PROGRAM OtherDevice_外部機器
VAR
    FH_M : BOOL;
    GT2_M : BOOL;
    IAI_M : BOOL;
    HMI_M : BOOL;
    FH_A_ST1_M : ARRAY[0..99] OF Bool;  (* [1] ST1 FH測定中; [5] ST1 測定完了 *)
    FH_A_ST1_OK : BOOL;  (* ST1 OK判定 *)
    FH_A_ST1_NG : BOOL;  (* ST1 NG 判定 *)
    FH_A_ST1_TON : ARRAY[0..99] OF TON;
    FH_A_ST1_TOF : ARRAY[0..99] OF TOF;
    ４ : UINT;
    ConvWordIndex : INT;  (* ワード処理ループの添字。（2台を順番に処理する作業用。運転指令は入れない） *)
    ConvAxisIndex : INT;  (* 軸処理ループの添字1～6。（2台を順番に処理する作業用。運転指令は入れない） *)
    ConvBase : INT;  (* 軸データの先頭添字8/16/24/32/40/48。（2台を順番に処理する作業用。運転指令は入れない） *)
    ConvDWord : DWORD;  (* 32bitの分割・結合に使うビット列。（2台を順番に処理する作業用。運転指令は入れない） *)
    ConvPos : DINT;  (* 0.01mm単位の符号付き目標位置。（2台を順番に処理する作業用。運転指令は入れない） *)
    ConvBand : UDINT;  (* 0.01mm単位の非負位置決め幅（内部推奨型）。（2台を順番に処理する作業用。運転指令は入れない） *)
    ConvSpeed : UINT;  (* 速度の送信整数。（2台を順番に処理する作業用。運転指令は入れない） *)
    ConvAccDec : UINT;  (* 加減速度の送信整数。（2台を順番に処理する作業用。運転指令は入れない） *)
    ConvPush : UINT;  (* 押付け電流制限の送信整数。（2台を順番に処理する作業用。運転指令は入れない） *)
    ConvScaled : LREAL;  (* 単位換算の作業値。（2台を順番に処理する作業用。運転指令は入れない） *)
    ConvWord : WORD;  (* バイト交換の作業ワード。（2台を順番に処理する作業用。運転指令は入れない） *)
    ConvUnitOK : BOOL;  (* 速度単位が1.0または0.1であること。（2台を順番に処理する作業用。運転指令は入れない） *)
END_VAR
VAR_EXTERNAL
    HMI_MessageNo : ARRAY[0..9] OF UINT;
    HMI_Message : ARRAY[0..9] OF String[256];
    HMI_Language : BOOL;
    FH_Line0_Trigger_Ready_1 : BOOL;
    FH_Line0_Trigger_1 : BOOL;
    M9999 : BOOL;
    FH_Line0_Busy_1 : BOOL;
    FH_Line0_Result_Notification_1 : BOOL;
    FH_Line0_DINT_Result_Data_0_1 : DINT;
    FH_Line0_DINT_Result_Data_1_1 : DINT;
    FH_Line0_DINT_Result_Data_2_1 : DINT;
    FH_Line0_Command_Code_1 : DWORD;
    FH_Line0_Command_Request_1 : BOOL;
    FH_Line0_Command_Completion_1 : BOOL;
    MdlChg : BOOL;  (* 機種切替：ON【GA120】 OFF【GA90】 *)
    FH_Line0_Error_Status_1 : BOOL;
    FH_5552_10_A_Auto : BOOL;  (* ST1 FH測定開始 *)
    FH_A_ST1_Manual : BOOL;  (* ST1 *)
    Pause : ARRAY[0..99] OF Bool;
    FH_A_ST1_Done : BOOL;  (* ST1 画像検査完了 *)
    Station_A_Data : ARRAY[0..8] OF sData;
    DLEP1_OUT : ARRAY[0..79] OF BOOL;
    DLEP2_OUT : ARRAY[0..79] OF BOOL;
    DLEP1_IN : ARRAY[0..167] OF byte;
    DLEP2_IN : ARRAY[0..167] OF byte;
    DLEP2_IN_Error : BOOL;  (* B(右側)センサエラー *)
    DLEP1_IN_Error : BOOL;  (* A(右側)センサエラー *)
    GT2_A_CurrentVal : INT;  (* A(左側) 測定値 *)
    GT2_B_CurrentVal : INT;  (* B(右側) 測定値 *)
    Hgt_A_Ins_Data : LREAL;  (* A測定データに変換 *)
    Hgt_B_Ins_Data : LREAL;
    Hgt_A_ComputedValueData : LREAL;  (* A測定データ+13.000mm 算定データ *)
    Hgt_B_ComputedValueData : LREAL;  (* B測定データ+13.000mm 算定データ *)
    E001_In_IN00_2004_01 : UINT;  (* RCON1（Node1） RCON→PLC 【IN00】共通 ゲートウェイ状態信号0 *)
    E001_In_IN01_2004_02 : UINT;  (* RCON1（Node1） RCON→PLC 【IN01】共通 ゲートウェイ状態信号1（軸No.0～15リンク状態） *)
    E001_In_IN02_2004_03 : UINT;  (* RCON1（Node1） RCON→PLC 【IN02】共通 電源ユニット状態信号0 *)
    E001_In_IN03_2004_04 : UINT;  (* RCON1（Node1） RCON→PLC 【IN03】共通 電源ユニット状態信号1 *)
    E001_In_IN04_2004_05 : UINT;  (* RCON1（Node1） RCON→PLC 【IN04】共通 電源ユニット状態信号2 *)
    E001_In_IN05_2004_06 : UINT;  (* RCON1（Node1） RCON→PLC 【IN05】共通 電源ユニット状態信号3 *)
    E001_In_IN06_2004_07 : UINT;  (* RCON1（Node1） RCON→PLC 【IN06】共通 電源ユニット状態信号4／軽故障メンテナンス（設定依存） *)
    E001_In_IN07_2004_08 : UINT;  (* RCON1（Node1） RCON→PLC 【IN07】共通 共通予約領域（使用禁止・占有あり） *)
    E001_In_IN08_2004_09 : UINT;  (* RCON1（Node1） RCON→PLC 【IN08】1軸目（No.0） 現在位置 下位ワード *)
    E001_In_IN09_2004_0A : UINT;  (* RCON1（Node1） RCON→PLC 【IN09】1軸目（No.0） 現在位置 上位ワード *)
    E001_In_IN10_2004_0B : UINT;  (* RCON1（Node1） RCON→PLC 【IN10】1軸目（No.0） 現在電流 下位ワード（PCは指令電流） *)
    E001_In_IN11_2004_0C : UINT;  (* RCON1（Node1） RCON→PLC 【IN11】1軸目（No.0） 現在電流 上位ワード（PCは指令電流） *)
    E001_In_IN12_2004_0D : UINT;  (* RCON1（Node1） RCON→PLC 【IN12】1軸目（No.0） 現在速度（負方向は2の補数） *)
    E001_In_IN13_2004_0E : UINT;  (* RCON1（Node1） RCON→PLC 【IN13】1軸目（No.0） 予約領域（使用禁止） *)
    E001_In_IN14_2004_0F : UINT;  (* RCON1（Node1） RCON→PLC 【IN14】1軸目（No.0） アラームコード（簡易コードではない） *)
    E001_In_IN15_2004_10 : UINT;  (* RCON1（Node1） RCON→PLC 【IN15】1軸目（No.0） 軸状態信号（PEND・SV等） *)
    E001_In_IN16_2004_11 : UINT;  (* RCON1（Node1） RCON→PLC 【IN16】2軸目（No.1） 現在位置 下位ワード *)
    E001_In_IN17_2004_12 : UINT;  (* RCON1（Node1） RCON→PLC 【IN17】2軸目（No.1） 現在位置 上位ワード *)
    E001_In_IN18_2004_13 : UINT;  (* RCON1（Node1） RCON→PLC 【IN18】2軸目（No.1） 現在電流 下位ワード（PCは指令電流） *)
    E001_In_IN19_2004_14 : UINT;  (* RCON1（Node1） RCON→PLC 【IN19】2軸目（No.1） 現在電流 上位ワード（PCは指令電流） *)
    E001_In_IN20_2004_15 : UINT;  (* RCON1（Node1） RCON→PLC 【IN20】2軸目（No.1） 現在速度（負方向は2の補数） *)
    E001_In_IN21_2004_16 : UINT;  (* RCON1（Node1） RCON→PLC 【IN21】2軸目（No.1） 予約領域（使用禁止） *)
    E001_In_IN22_2004_17 : UINT;  (* RCON1（Node1） RCON→PLC 【IN22】2軸目（No.1） アラームコード（簡易コードではない） *)
    E001_In_IN23_2004_18 : UINT;  (* RCON1（Node1） RCON→PLC 【IN23】2軸目（No.1） 軸状態信号（PEND・SV等） *)
    E001_In_IN24_2004_19 : UINT;  (* RCON1（Node1） RCON→PLC 【IN24】3軸目（No.2） 現在位置 下位ワード *)
    E001_In_IN25_2004_1A : UINT;  (* RCON1（Node1） RCON→PLC 【IN25】3軸目（No.2） 現在位置 上位ワード *)
    E001_In_IN26_2004_1B : UINT;  (* RCON1（Node1） RCON→PLC 【IN26】3軸目（No.2） 現在電流 下位ワード（PCは指令電流） *)
    E001_In_IN27_2004_1C : UINT;  (* RCON1（Node1） RCON→PLC 【IN27】3軸目（No.2） 現在電流 上位ワード（PCは指令電流） *)
    E001_In_IN28_2004_1D : UINT;  (* RCON1（Node1） RCON→PLC 【IN28】3軸目（No.2） 現在速度（負方向は2の補数） *)
    E001_In_IN29_2004_1E : UINT;  (* RCON1（Node1） RCON→PLC 【IN29】3軸目（No.2） 予約領域（使用禁止） *)
    E001_In_IN30_2004_1F : UINT;  (* RCON1（Node1） RCON→PLC 【IN30】3軸目（No.2） アラームコード（簡易コードではない） *)
    E001_In_IN31_2004_20 : UINT;  (* RCON1（Node1） RCON→PLC 【IN31】3軸目（No.2） 軸状態信号（PEND・SV等） *)
    E001_In_IN32_2004_21 : UINT;  (* RCON1（Node1） RCON→PLC 【IN32】4軸目（No.3） 現在位置 下位ワード *)
    E001_In_IN33_2004_22 : UINT;  (* RCON1（Node1） RCON→PLC 【IN33】4軸目（No.3） 現在位置 上位ワード *)
    E001_In_IN34_2004_23 : UINT;  (* RCON1（Node1） RCON→PLC 【IN34】4軸目（No.3） 現在電流 下位ワード（PCは指令電流） *)
    E001_In_IN35_2004_24 : UINT;  (* RCON1（Node1） RCON→PLC 【IN35】4軸目（No.3） 現在電流 上位ワード（PCは指令電流） *)
    E001_In_IN36_2004_25 : UINT;  (* RCON1（Node1） RCON→PLC 【IN36】4軸目（No.3） 現在速度（負方向は2の補数） *)
    E001_In_IN37_2004_26 : UINT;  (* RCON1（Node1） RCON→PLC 【IN37】4軸目（No.3） 予約領域（使用禁止） *)
    E001_In_IN38_2004_27 : UINT;  (* RCON1（Node1） RCON→PLC 【IN38】4軸目（No.3） アラームコード（簡易コードではない） *)
    E001_In_IN39_2004_28 : UINT;  (* RCON1（Node1） RCON→PLC 【IN39】4軸目（No.3） 軸状態信号（PEND・SV等） *)
    E001_In_IN40_2004_29 : UINT;  (* RCON1（Node1） RCON→PLC 【IN40】5軸目（No.4） 現在位置 下位ワード *)
    E001_In_IN41_2004_2A : UINT;  (* RCON1（Node1） RCON→PLC 【IN41】5軸目（No.4） 現在位置 上位ワード *)
    E001_In_IN42_2004_2B : UINT;  (* RCON1（Node1） RCON→PLC 【IN42】5軸目（No.4） 現在電流 下位ワード（PCは指令電流） *)
    E001_In_IN43_2004_2C : UINT;  (* RCON1（Node1） RCON→PLC 【IN43】5軸目（No.4） 現在電流 上位ワード（PCは指令電流） *)
    E001_In_IN44_2004_2D : UINT;  (* RCON1（Node1） RCON→PLC 【IN44】5軸目（No.4） 現在速度（負方向は2の補数） *)
    E001_In_IN45_2004_2E : UINT;  (* RCON1（Node1） RCON→PLC 【IN45】5軸目（No.4） 予約領域（使用禁止） *)
    E001_In_IN46_2004_2F : UINT;  (* RCON1（Node1） RCON→PLC 【IN46】5軸目（No.4） アラームコード（簡易コードではない） *)
    E001_In_IN47_2004_30 : UINT;  (* RCON1（Node1） RCON→PLC 【IN47】5軸目（No.4） 軸状態信号（PEND・SV等） *)
    E001_In_IN48_2004_31 : UINT;  (* RCON1（Node1） RCON→PLC 【IN48】6軸目（No.5） 現在位置 下位ワード *)
    E001_In_IN49_2004_32 : UINT;  (* RCON1（Node1） RCON→PLC 【IN49】6軸目（No.5） 現在位置 上位ワード *)
    E001_In_IN50_2004_33 : UINT;  (* RCON1（Node1） RCON→PLC 【IN50】6軸目（No.5） 現在電流 下位ワード（PCは指令電流） *)
    E001_In_IN51_2004_34 : UINT;  (* RCON1（Node1） RCON→PLC 【IN51】6軸目（No.5） 現在電流 上位ワード（PCは指令電流） *)
    E001_In_IN52_2004_35 : UINT;  (* RCON1（Node1） RCON→PLC 【IN52】6軸目（No.5） 現在速度（負方向は2の補数） *)
    E001_In_IN53_2004_36 : UINT;  (* RCON1（Node1） RCON→PLC 【IN53】6軸目（No.5） 予約領域（使用禁止） *)
    E001_In_IN54_2004_37 : UINT;  (* RCON1（Node1） RCON→PLC 【IN54】6軸目（No.5） アラームコード（簡易コードではない） *)
    E001_In_IN55_2004_38 : UINT;  (* RCON1（Node1） RCON→PLC 【IN55】6軸目（No.5） 軸状態信号（PEND・SV等） *)
    E001_In_IN56_2004_39 : UINT;  (* RCON1（Node1） 【IN56】用途未確認領域。今回の軸データ変換では未使用。 *)
    E001_In_IN57_2004_3A : UINT;  (* RCON1（Node1） 【IN57】用途未確認領域。今回の軸データ変換では未使用。 *)
    E001_In_IN58_2004_3B : UINT;  (* RCON1（Node1） 【IN58】用途未確認領域。今回の軸データ変換では未使用。 *)
    E001_In_IN59_2004_3C : UINT;  (* RCON1（Node1） 【IN59】用途未確認領域。今回の軸データ変換では未使用。 *)
    E001_In_IN60_2004_3D : UINT;  (* RCON1（Node1） 【IN60】用途未確認領域。今回の軸データ変換では未使用。 *)
    E001_In_IN61_2004_3E : UINT;  (* RCON1（Node1） 【IN61】用途未確認領域。今回の軸データ変換では未使用。 *)
    E001_In_IN62_2004_3F : UINT;  (* RCON1（Node1） 【IN62】用途未確認領域。今回の軸データ変換では未使用。 *)
    E001_In_IN63_2004_40 : UINT;  (* RCON1（Node1） 【IN63】用途未確認領域。今回の軸データ変換では未使用。 *)
    E001_In_IN64_2004_41 : UINT;  (* RCON1（Node1） 【IN64】用途未確認領域。今回の軸データ変換では未使用。 *)
    E001_In_IN65_2004_42 : UINT;  (* RCON1（Node1） 【IN65】用途未確認領域。今回の軸データ変換では未使用。 *)
    E001_In_IN66_2004_43 : UINT;  (* RCON1（Node1） 【IN66】用途未確認領域。今回の軸データ変換では未使用。 *)
    E001_In_IN67_2004_44 : UINT;  (* RCON1（Node1） 【IN67】用途未確認領域。今回の軸データ変換では未使用。 *)
    E001_In_IN68_2004_45 : UINT;  (* RCON1（Node1） 【IN68】用途未確認領域。今回の軸データ変換では未使用。 *)
    E001_In_IN69_2004_46 : UINT;  (* RCON1（Node1） 【IN69】用途未確認領域。今回の軸データ変換では未使用。 *)
    E001_In_IN70_2004_47 : UINT;  (* RCON1（Node1） 【IN70】用途未確認領域。今回の軸データ変換では未使用。 *)
    E001_In_IN71_2004_48 : UINT;  (* RCON1（Node1） 【IN71】用途未確認領域。今回の軸データ変換では未使用。 *)
    E001_Out_OUT00_2003_01 : UINT;  (* RCON1（Node1） PLC→RCON 【OUT00】共通 ゲートウェイ制御信号0（MON等） *)
    E001_Out_OUT08_2003_09 : UINT;  (* RCON1（Node1） PLC→RCON 【OUT08】1軸目（No.0） 目標位置 下位ワード *)
    E001_Out_OUT09_2003_0A : UINT;  (* RCON1（Node1） PLC→RCON 【OUT09】1軸目（No.0） 目標位置 上位ワード *)
    E001_Out_OUT10_2003_0B : UINT;  (* RCON1（Node1） PLC→RCON 【OUT10】1軸目（No.0） 位置決め幅 下位ワード *)
    E001_Out_OUT11_2003_0C : UINT;  (* RCON1（Node1） PLC→RCON 【OUT11】1軸目（No.0） 位置決め幅 上位ワード *)
    E001_Out_OUT12_2003_0D : UINT;  (* RCON1（Node1） PLC→RCON 【OUT12】1軸目（No.0） 速度指令 *)
    E001_Out_OUT13_2003_0E : UINT;  (* RCON1（Node1） PLC→RCON 【OUT13】1軸目（No.0） 加減速度指令（加速・減速共通） *)
    E001_Out_OUT14_2003_0F : UINT;  (* RCON1（Node1） PLC→RCON 【OUT14】1軸目（No.0） 押付け電流制限値 *)
    E001_Out_OUT15_2003_10 : UINT;  (* RCON1（Node1） PLC→RCON 【OUT15】1軸目（No.0） 軸制御信号（DSTR・SON等） *)
    E001_Out_OUT16_2003_11 : UINT;  (* RCON1（Node1） PLC→RCON 【OUT16】2軸目（No.1） 目標位置 下位ワード *)
    E001_Out_OUT17_2003_12 : UINT;  (* RCON1（Node1） PLC→RCON 【OUT17】2軸目（No.1） 目標位置 上位ワード *)
    E001_Out_OUT18_2003_13 : UINT;  (* RCON1（Node1） PLC→RCON 【OUT18】2軸目（No.1） 位置決め幅 下位ワード *)
    E001_Out_OUT19_2003_14 : UINT;  (* RCON1（Node1） PLC→RCON 【OUT19】2軸目（No.1） 位置決め幅 上位ワード *)
    E001_Out_OUT20_2003_15 : UINT;  (* RCON1（Node1） PLC→RCON 【OUT20】2軸目（No.1） 速度指令 *)
    E001_Out_OUT21_2003_16 : UINT;  (* RCON1（Node1） PLC→RCON 【OUT21】2軸目（No.1） 加減速度指令（加速・減速共通） *)
    E001_Out_OUT22_2003_17 : UINT;  (* RCON1（Node1） PLC→RCON 【OUT22】2軸目（No.1） 押付け電流制限値 *)
    E001_Out_OUT23_2003_18 : UINT;  (* RCON1（Node1） PLC→RCON 【OUT23】2軸目（No.1） 軸制御信号（DSTR・SON等） *)
    E001_Out_OUT24_2003_19 : UINT;  (* RCON1（Node1） PLC→RCON 【OUT24】3軸目（No.2） 目標位置 下位ワード *)
    E001_Out_OUT25_2003_1A : UINT;  (* RCON1（Node1） PLC→RCON 【OUT25】3軸目（No.2） 目標位置 上位ワード *)
    E001_Out_OUT26_2003_1B : UINT;  (* RCON1（Node1） PLC→RCON 【OUT26】3軸目（No.2） 位置決め幅 下位ワード *)
    E001_Out_OUT27_2003_1C : UINT;  (* RCON1（Node1） PLC→RCON 【OUT27】3軸目（No.2） 位置決め幅 上位ワード *)
    E001_Out_OUT28_2003_1D : UINT;  (* RCON1（Node1） PLC→RCON 【OUT28】3軸目（No.2） 速度指令 *)
    E001_Out_OUT29_2003_1E : UINT;  (* RCON1（Node1） PLC→RCON 【OUT29】3軸目（No.2） 加減速度指令（加速・減速共通） *)
    E001_Out_OUT30_2003_1F : UINT;  (* RCON1（Node1） PLC→RCON 【OUT30】3軸目（No.2） 押付け電流制限値 *)
    E001_Out_OUT31_2003_20 : UINT;  (* RCON1（Node1） PLC→RCON 【OUT31】3軸目（No.2） 軸制御信号（DSTR・SON等） *)
    E001_Out_OUT32_2003_21 : UINT;  (* RCON1（Node1） PLC→RCON 【OUT32】4軸目（No.3） 目標位置 下位ワード *)
    E001_Out_OUT33_2003_22 : UINT;  (* RCON1（Node1） PLC→RCON 【OUT33】4軸目（No.3） 目標位置 上位ワード *)
    E001_Out_OUT34_2003_23 : UINT;  (* RCON1（Node1） PLC→RCON 【OUT34】4軸目（No.3） 位置決め幅 下位ワード *)
    E001_Out_OUT35_2003_24 : UINT;  (* RCON1（Node1） PLC→RCON 【OUT35】4軸目（No.3） 位置決め幅 上位ワード *)
    E001_Out_OUT36_2003_25 : UINT;  (* RCON1（Node1） PLC→RCON 【OUT36】4軸目（No.3） 速度指令 *)
    E001_Out_OUT37_2003_26 : UINT;  (* RCON1（Node1） PLC→RCON 【OUT37】4軸目（No.3） 加減速度指令（加速・減速共通） *)
    E001_Out_OUT38_2003_27 : UINT;  (* RCON1（Node1） PLC→RCON 【OUT38】4軸目（No.3） 押付け電流制限値 *)
    E001_Out_OUT39_2003_28 : UINT;  (* RCON1（Node1） PLC→RCON 【OUT39】4軸目（No.3） 軸制御信号（DSTR・SON等） *)
    E001_Out_OUT40_2003_29 : UINT;  (* RCON1（Node1） PLC→RCON 【OUT40】5軸目（No.4） 目標位置 下位ワード *)
    E001_Out_OUT41_2003_2A : UINT;  (* RCON1（Node1） PLC→RCON 【OUT41】5軸目（No.4） 目標位置 上位ワード *)
    E001_Out_OUT42_2003_2B : UINT;  (* RCON1（Node1） PLC→RCON 【OUT42】5軸目（No.4） 位置決め幅 下位ワード *)
    E001_Out_OUT43_2003_2C : UINT;  (* RCON1（Node1） PLC→RCON 【OUT43】5軸目（No.4） 位置決め幅 上位ワード *)
    E001_Out_OUT44_2003_2D : UINT;  (* RCON1（Node1） PLC→RCON 【OUT44】5軸目（No.4） 速度指令 *)
    E001_Out_OUT45_2003_2E : UINT;  (* RCON1（Node1） PLC→RCON 【OUT45】5軸目（No.4） 加減速度指令（加速・減速共通） *)
    E001_Out_OUT46_2003_2F : UINT;  (* RCON1（Node1） PLC→RCON 【OUT46】5軸目（No.4） 押付け電流制限値 *)
    E001_Out_OUT47_2003_30 : UINT;  (* RCON1（Node1） PLC→RCON 【OUT47】5軸目（No.4） 軸制御信号（DSTR・SON等） *)
    E001_Out_OUT48_2003_31 : UINT;  (* RCON1（Node1） PLC→RCON 【OUT48】6軸目（No.5） 目標位置 下位ワード *)
    E001_Out_OUT49_2003_32 : UINT;  (* RCON1（Node1） PLC→RCON 【OUT49】6軸目（No.5） 目標位置 上位ワード *)
    E001_Out_OUT50_2003_33 : UINT;  (* RCON1（Node1） PLC→RCON 【OUT50】6軸目（No.5） 位置決め幅 下位ワード *)
    E001_Out_OUT51_2003_34 : UINT;  (* RCON1（Node1） PLC→RCON 【OUT51】6軸目（No.5） 位置決め幅 上位ワード *)
    E001_Out_OUT52_2003_35 : UINT;  (* RCON1（Node1） PLC→RCON 【OUT52】6軸目（No.5） 速度指令 *)
    E001_Out_OUT53_2003_36 : UINT;  (* RCON1（Node1） PLC→RCON 【OUT53】6軸目（No.5） 加減速度指令（加速・減速共通） *)
    E001_Out_OUT54_2003_37 : UINT;  (* RCON1（Node1） PLC→RCON 【OUT54】6軸目（No.5） 押付け電流制限値 *)
    E001_Out_OUT55_2003_38 : UINT;  (* RCON1（Node1） PLC→RCON 【OUT55】6軸目（No.5） 軸制御信号（DSTR・SON等） *)
    E005_In_IN00_2004_01_1 : UINT;  (* RCON2（Node5） RCON→PLC 【IN00】共通 ゲートウェイ状態信号0 *)
    E005_In_IN01_2004_02_1 : UINT;  (* RCON2（Node5） RCON→PLC 【IN01】共通 ゲートウェイ状態信号1（軸No.0～15リンク状態） *)
    E005_In_IN02_2004_03_1 : UINT;  (* RCON2（Node5） RCON→PLC 【IN02】共通 電源ユニット状態信号0 *)
    E005_In_IN03_2004_04_1 : UINT;  (* RCON2（Node5） RCON→PLC 【IN03】共通 電源ユニット状態信号1 *)
    E005_In_IN04_2004_05_1 : UINT;  (* RCON2（Node5） RCON→PLC 【IN04】共通 電源ユニット状態信号2 *)
    E005_In_IN05_2004_06_1 : UINT;  (* RCON2（Node5） RCON→PLC 【IN05】共通 電源ユニット状態信号3 *)
    E005_In_IN06_2004_07_1 : UINT;  (* RCON2（Node5） RCON→PLC 【IN06】共通 電源ユニット状態信号4／軽故障メンテナンス（設定依存） *)
    E005_In_IN07_2004_08_1 : UINT;  (* RCON2（Node5） RCON→PLC 【IN07】共通 共通予約領域（使用禁止・占有あり） *)
    E005_In_IN08_2004_09_1 : UINT;  (* RCON2（Node5） RCON→PLC 【IN08】1軸目（No.0） 現在位置 下位ワード *)
    E005_In_IN09_2004_0A_1 : UINT;  (* RCON2（Node5） RCON→PLC 【IN09】1軸目（No.0） 現在位置 上位ワード *)
    E005_In_IN10_2004_0B_1 : UINT;  (* RCON2（Node5） RCON→PLC 【IN10】1軸目（No.0） 現在電流 下位ワード（PCは指令電流） *)
    E005_In_IN11_2004_0C_1 : UINT;  (* RCON2（Node5） RCON→PLC 【IN11】1軸目（No.0） 現在電流 上位ワード（PCは指令電流） *)
    E005_In_IN12_2004_0D_1 : UINT;  (* RCON2（Node5） RCON→PLC 【IN12】1軸目（No.0） 現在速度（負方向は2の補数） *)
    E005_In_IN13_2004_0E_1 : UINT;  (* RCON2（Node5） RCON→PLC 【IN13】1軸目（No.0） 予約領域（使用禁止） *)
    E005_In_IN14_2004_0F_1 : UINT;  (* RCON2（Node5） RCON→PLC 【IN14】1軸目（No.0） アラームコード（簡易コードではない） *)
    E005_In_IN15_2004_10_1 : UINT;  (* RCON2（Node5） RCON→PLC 【IN15】1軸目（No.0） 軸状態信号（PEND・SV等） *)
    E005_In_IN16_2004_11_1 : UINT;  (* RCON2（Node5） RCON→PLC 【IN16】2軸目（No.1） 現在位置 下位ワード *)
    E005_In_IN17_2004_12_1 : UINT;  (* RCON2（Node5） RCON→PLC 【IN17】2軸目（No.1） 現在位置 上位ワード *)
    E005_In_IN18_2004_13_1 : UINT;  (* RCON2（Node5） RCON→PLC 【IN18】2軸目（No.1） 現在電流 下位ワード（PCは指令電流） *)
    E005_In_IN19_2004_14_1 : UINT;  (* RCON2（Node5） RCON→PLC 【IN19】2軸目（No.1） 現在電流 上位ワード（PCは指令電流） *)
    E005_In_IN20_2004_15_1 : UINT;  (* RCON2（Node5） RCON→PLC 【IN20】2軸目（No.1） 現在速度（負方向は2の補数） *)
    E005_In_IN21_2004_16_1 : UINT;  (* RCON2（Node5） RCON→PLC 【IN21】2軸目（No.1） 予約領域（使用禁止） *)
    E005_In_IN22_2004_17_1 : UINT;  (* RCON2（Node5） RCON→PLC 【IN22】2軸目（No.1） アラームコード（簡易コードではない） *)
    E005_In_IN23_2004_18_1 : UINT;  (* RCON2（Node5） RCON→PLC 【IN23】2軸目（No.1） 軸状態信号（PEND・SV等） *)
    E005_In_IN24_2004_19_1 : UINT;  (* RCON2（Node5） RCON→PLC 【IN24】3軸目（No.2） 現在位置 下位ワード *)
    E005_In_IN25_2004_1A_1 : UINT;  (* RCON2（Node5） RCON→PLC 【IN25】3軸目（No.2） 現在位置 上位ワード *)
    E005_In_IN26_2004_1B_1 : UINT;  (* RCON2（Node5） RCON→PLC 【IN26】3軸目（No.2） 現在電流 下位ワード（PCは指令電流） *)
    E005_In_IN27_2004_1C_1 : UINT;  (* RCON2（Node5） RCON→PLC 【IN27】3軸目（No.2） 現在電流 上位ワード（PCは指令電流） *)
    E005_In_IN28_2004_1D_1 : UINT;  (* RCON2（Node5） RCON→PLC 【IN28】3軸目（No.2） 現在速度（負方向は2の補数） *)
    E005_In_IN29_2004_1E_1 : UINT;  (* RCON2（Node5） RCON→PLC 【IN29】3軸目（No.2） 予約領域（使用禁止） *)
    E005_In_IN30_2004_1F_1 : UINT;  (* RCON2（Node5） RCON→PLC 【IN30】3軸目（No.2） アラームコード（簡易コードではない） *)
    E005_In_IN31_2004_20_1 : UINT;  (* RCON2（Node5） RCON→PLC 【IN31】3軸目（No.2） 軸状態信号（PEND・SV等） *)
    E005_In_IN32_2004_21_1 : UINT;  (* RCON2（Node5） RCON→PLC 【IN32】4軸目（No.3） 現在位置 下位ワード *)
    E005_In_IN33_2004_22_1 : UINT;  (* RCON2（Node5） RCON→PLC 【IN33】4軸目（No.3） 現在位置 上位ワード *)
    E005_In_IN34_2004_23_1 : UINT;  (* RCON2（Node5） RCON→PLC 【IN34】4軸目（No.3） 現在電流 下位ワード（PCは指令電流） *)
    E005_In_IN35_2004_24_1 : UINT;  (* RCON2（Node5） RCON→PLC 【IN35】4軸目（No.3） 現在電流 上位ワード（PCは指令電流） *)
    E005_In_IN36_2004_25_1 : UINT;  (* RCON2（Node5） RCON→PLC 【IN36】4軸目（No.3） 現在速度（負方向は2の補数） *)
    E005_In_IN37_2004_26_1 : UINT;  (* RCON2（Node5） RCON→PLC 【IN37】4軸目（No.3） 予約領域（使用禁止） *)
    E005_In_IN38_2004_27_1 : UINT;  (* RCON2（Node5） RCON→PLC 【IN38】4軸目（No.3） アラームコード（簡易コードではない） *)
    E005_In_IN39_2004_28_1 : UINT;  (* RCON2（Node5） RCON→PLC 【IN39】4軸目（No.3） 軸状態信号（PEND・SV等） *)
    E005_In_IN40_2004_29_1 : UINT;  (* RCON2（Node5） RCON→PLC 【IN40】5軸目（No.4） 現在位置 下位ワード *)
    E005_In_IN41_2004_2A_1 : UINT;  (* RCON2（Node5） RCON→PLC 【IN41】5軸目（No.4） 現在位置 上位ワード *)
    E005_In_IN42_2004_2B_1 : UINT;  (* RCON2（Node5） RCON→PLC 【IN42】5軸目（No.4） 現在電流 下位ワード（PCは指令電流） *)
    E005_In_IN43_2004_2C_1 : UINT;  (* RCON2（Node5） RCON→PLC 【IN43】5軸目（No.4） 現在電流 上位ワード（PCは指令電流） *)
    E005_In_IN44_2004_2D_1 : UINT;  (* RCON2（Node5） RCON→PLC 【IN44】5軸目（No.4） 現在速度（負方向は2の補数） *)
    E005_In_IN45_2004_2E_1 : UINT;  (* RCON2（Node5） RCON→PLC 【IN45】5軸目（No.4） 予約領域（使用禁止） *)
    E005_In_IN46_2004_2F_1 : UINT;  (* RCON2（Node5） RCON→PLC 【IN46】5軸目（No.4） アラームコード（簡易コードではない） *)
    E005_In_IN47_2004_30_1 : UINT;  (* RCON2（Node5） RCON→PLC 【IN47】5軸目（No.4） 軸状態信号（PEND・SV等） *)
    E005_In_IN48_2004_31_1 : UINT;  (* RCON2（Node5） 【IN48】用途未確認領域。今回の軸データ変換では未使用。 *)
    E005_In_IN49_2004_32_1 : UINT;  (* RCON2（Node5） 【IN49】用途未確認領域。今回の軸データ変換では未使用。 *)
    E005_In_IN50_2004_33_1 : UINT;  (* RCON2（Node5） 【IN50】用途未確認領域。今回の軸データ変換では未使用。 *)
    E005_In_IN51_2004_34_1 : UINT;  (* RCON2（Node5） 【IN51】用途未確認領域。今回の軸データ変換では未使用。 *)
    E005_In_IN52_2004_35_1 : UINT;  (* RCON2（Node5） 【IN52】用途未確認領域。今回の軸データ変換では未使用。 *)
    E005_In_IN53_2004_36_1 : UINT;  (* RCON2（Node5） 【IN53】用途未確認領域。今回の軸データ変換では未使用。 *)
    E005_In_IN54_2004_37_1 : UINT;  (* RCON2（Node5） 【IN54】用途未確認領域。今回の軸データ変換では未使用。 *)
    E005_In_IN55_2004_38_1 : UINT;  (* RCON2（Node5） 【IN55】用途未確認領域。今回の軸データ変換では未使用。 *)
    E005_Out_OUT00_2003_01_1 : UINT;  (* RCON2（Node5） PLC→RCON 【OUT00】共通 ゲートウェイ制御信号0（MON等） *)
    E005_Out_OUT08_2003_09_1 : UINT;  (* RCON2（Node5） PLC→RCON 【OUT08】1軸目（No.0） 目標位置 下位ワード *)
    E005_Out_OUT09_2003_0A_1 : UINT;  (* RCON2（Node5） PLC→RCON 【OUT09】1軸目（No.0） 目標位置 上位ワード *)
    E005_Out_OUT10_2003_0B_1 : UINT;  (* RCON2（Node5） PLC→RCON 【OUT10】1軸目（No.0） 位置決め幅 下位ワード *)
    E005_Out_OUT11_2003_0C_1 : UINT;  (* RCON2（Node5） PLC→RCON 【OUT11】1軸目（No.0） 位置決め幅 上位ワード *)
    E005_Out_OUT12_2003_0D_1 : UINT;  (* RCON2（Node5） PLC→RCON 【OUT12】1軸目（No.0） 速度指令 *)
    E005_Out_OUT13_2003_0E_1 : UINT;  (* RCON2（Node5） PLC→RCON 【OUT13】1軸目（No.0） 加減速度指令（加速・減速共通） *)
    E005_Out_OUT14_2003_0F_1 : UINT;  (* RCON2（Node5） PLC→RCON 【OUT14】1軸目（No.0） 押付け電流制限値 *)
    E005_Out_OUT15_2003_10_1 : UINT;  (* RCON2（Node5） PLC→RCON 【OUT15】1軸目（No.0） 軸制御信号（DSTR・SON等） *)
    E005_Out_OUT16_2003_11_1 : UINT;  (* RCON2（Node5） PLC→RCON 【OUT16】2軸目（No.1） 目標位置 下位ワード *)
    E005_Out_OUT17_2003_12_1 : UINT;  (* RCON2（Node5） PLC→RCON 【OUT17】2軸目（No.1） 目標位置 上位ワード *)
    E005_Out_OUT18_2003_13_1 : UINT;  (* RCON2（Node5） PLC→RCON 【OUT18】2軸目（No.1） 位置決め幅 下位ワード *)
    E005_Out_OUT19_2003_14_1 : UINT;  (* RCON2（Node5） PLC→RCON 【OUT19】2軸目（No.1） 位置決め幅 上位ワード *)
    E005_Out_OUT20_2003_15_1 : UINT;  (* RCON2（Node5） PLC→RCON 【OUT20】2軸目（No.1） 速度指令 *)
    E005_Out_OUT21_2003_16_1 : UINT;  (* RCON2（Node5） PLC→RCON 【OUT21】2軸目（No.1） 加減速度指令（加速・減速共通） *)
    E005_Out_OUT22_2003_17_1 : UINT;  (* RCON2（Node5） PLC→RCON 【OUT22】2軸目（No.1） 押付け電流制限値 *)
    E005_Out_OUT23_2003_18_1 : UINT;  (* RCON2（Node5） PLC→RCON 【OUT23】2軸目（No.1） 軸制御信号（DSTR・SON等） *)
    E005_Out_OUT24_2003_19_1 : UINT;  (* RCON2（Node5） PLC→RCON 【OUT24】3軸目（No.2） 目標位置 下位ワード *)
    E005_Out_OUT25_2003_1A_1 : UINT;  (* RCON2（Node5） PLC→RCON 【OUT25】3軸目（No.2） 目標位置 上位ワード *)
    E005_Out_OUT26_2003_1B_1 : UINT;  (* RCON2（Node5） PLC→RCON 【OUT26】3軸目（No.2） 位置決め幅 下位ワード *)
    E005_Out_OUT27_2003_1C_1 : UINT;  (* RCON2（Node5） PLC→RCON 【OUT27】3軸目（No.2） 位置決め幅 上位ワード *)
    E005_Out_OUT28_2003_1D_1 : UINT;  (* RCON2（Node5） PLC→RCON 【OUT28】3軸目（No.2） 速度指令 *)
    E005_Out_OUT29_2003_1E_1 : UINT;  (* RCON2（Node5） PLC→RCON 【OUT29】3軸目（No.2） 加減速度指令（加速・減速共通） *)
    E005_Out_OUT30_2003_1F_1 : UINT;  (* RCON2（Node5） PLC→RCON 【OUT30】3軸目（No.2） 押付け電流制限値 *)
    E005_Out_OUT31_2003_20_1 : UINT;  (* RCON2（Node5） PLC→RCON 【OUT31】3軸目（No.2） 軸制御信号（DSTR・SON等） *)
    E005_Out_OUT32_2003_21_1 : UINT;  (* RCON2（Node5） PLC→RCON 【OUT32】4軸目（No.3） 目標位置 下位ワード *)
    E005_Out_OUT33_2003_22_1 : UINT;  (* RCON2（Node5） PLC→RCON 【OUT33】4軸目（No.3） 目標位置 上位ワード *)
    E005_Out_OUT34_2003_23_1 : UINT;  (* RCON2（Node5） PLC→RCON 【OUT34】4軸目（No.3） 位置決め幅 下位ワード *)
    E005_Out_OUT35_2003_24_1 : UINT;  (* RCON2（Node5） PLC→RCON 【OUT35】4軸目（No.3） 位置決め幅 上位ワード *)
    E005_Out_OUT36_2003_25_1 : UINT;  (* RCON2（Node5） PLC→RCON 【OUT36】4軸目（No.3） 速度指令 *)
    E005_Out_OUT37_2003_26_1 : UINT;  (* RCON2（Node5） PLC→RCON 【OUT37】4軸目（No.3） 加減速度指令（加速・減速共通） *)
    E005_Out_OUT38_2003_27_1 : UINT;  (* RCON2（Node5） PLC→RCON 【OUT38】4軸目（No.3） 押付け電流制限値 *)
    E005_Out_OUT39_2003_28_1 : UINT;  (* RCON2（Node5） PLC→RCON 【OUT39】4軸目（No.3） 軸制御信号（DSTR・SON等） *)
    E005_Out_OUT40_2003_29_1 : UINT;  (* RCON2（Node5） PLC→RCON 【OUT40】5軸目（No.4） 目標位置 下位ワード *)
    E005_Out_OUT41_2003_2A_1 : UINT;  (* RCON2（Node5） PLC→RCON 【OUT41】5軸目（No.4） 目標位置 上位ワード *)
    E005_Out_OUT42_2003_2B_1 : UINT;  (* RCON2（Node5） PLC→RCON 【OUT42】5軸目（No.4） 位置決め幅 下位ワード *)
    E005_Out_OUT43_2003_2C_1 : UINT;  (* RCON2（Node5） PLC→RCON 【OUT43】5軸目（No.4） 位置決め幅 上位ワード *)
    E005_Out_OUT44_2003_2D_1 : UINT;  (* RCON2（Node5） PLC→RCON 【OUT44】5軸目（No.4） 速度指令 *)
    E005_Out_OUT45_2003_2E_1 : UINT;  (* RCON2（Node5） PLC→RCON 【OUT45】5軸目（No.4） 加減速度指令（加速・減速共通） *)
    E005_Out_OUT46_2003_2F_1 : UINT;  (* RCON2（Node5） PLC→RCON 【OUT46】5軸目（No.4） 押付け電流制限値 *)
    E005_Out_OUT47_2003_30_1 : UINT;  (* RCON2（Node5） PLC→RCON 【OUT47】5軸目（No.4） 軸制御信号（DSTR・SON等） *)
    RCON1_AxisApply : ARRAY[1..6] OF BOOL;  (* RCON1：初期FALSE。指定軸の8ワードを書込む。OFFは停止ではない。 *)
    RCON1_AxisLinked : ARRAY[1..6] OF BOOL;  (* RCON1：入力：軸No.0～5のリンク状態。 *)
    RCON1_AxisWritten : ARRAY[1..6] OF BOOL;  (* RCON1：各軸出力へ代入したサイクルのみTRUE。RCON受付・完了ではない。 *)
    RCON1_ByteOrderConfirmed : BOOL;  (* RCON1：初期FALSE。既知の位置とbitでワード順・バイト順を確認して設定。 *)
    RCON1_CommOK : BOOL;  (* RCON1：初期FALSE。CPUの実EtherCAT通信状態から別途作成。TRUE固定禁止。 *)
    RCON1_EncodeError : ARRAY[1..6] OF UINT;  (* RCON1：変換エラー番号。0正常、1単位、2位置、3幅、4速度、5加減速、6押付け、7両方向ジョグ。 *)
    RCON1_EncodeOK : ARRAY[1..6] OF BOOL;  (* RCON1：通信形式へ数値変換できたか。安全・運転許可ではない。 *)
    RCON1_GwAlarmCode : UINT;  (* RCON1：入力：ゲートウェイALMCの下位8bit。軸AlarmCodeとは別。 *)
    RCON1_GwApply : BOOL;  (* RCON1：初期FALSE。共通MON/RTEワードを書込む。 *)
    RCON1_GwAxisCommError : BOOL;  (* RCON1：入力：ゲートウェイと軸の通信異常ERRT。 *)
    RCON1_GwControllerCommLatch : BOOL;  (* RCON1：入力：運転中ERR-C保持LERC。 *)
    RCON1_GwHeavyAlarm : BOOL;  (* RCON1：入力：再起動が必要なゲートウェイ異常ALMH。 *)
    RCON1_GwLightAlarm : BOOL;  (* RCON1：入力：ゲートウェイ軽微異常ALML。 *)
    RCON1_GwMON_Request : BOOL;  (* RCON1：初期FALSE。ゲートウェイMON要求。論理b15。安全停止ではない。 *)
    RCON1_GwManual : BOOL;  (* RCON1：入力：MANUスイッチ選択MOD。 *)
    RCON1_GwRTE_Request : BOOL;  (* RCON1：初期FALSE。ゲートウェイ通信異常ラッチ解除要求。論理b13。 *)
    RCON1_GwRun : BOOL;  (* RCON1：入力：ゲートウェイ正常動作中RUN。 *)
    RCON1_GwSystemStop : BOOL;  (* RCON1：入力：システムSTOP入力による停止状態SEMG。安全回路の代用不可。 *)
    RCON1_GwWritten : BOOL;  (* RCON1：共通出力へ代入したサイクルのみTRUE。RCON受付の意味ではない。 *)
    RCON1_IN : ARRAY[1..6] OF ST_RCON_Direct_IN_Axis;  (* RCON1 6軸分 RCON→PLC 取得値・状態（内部変数・通信変換は別途） *)
    RCON1_LayoutConfirmed : BOOL;  (* RCON1：初期FALSE。全6軸直接数値指定・共通8W・軸順・占有を確認して設定。 *)
    RCON1_MotionPermit : ARRAY[1..6] OF BOOL;  (* RCON1：初期FALSE。機械範囲・安全・運転条件から別途作成する運転許可。単純TRUE固定禁止。 *)
    RCON1_OUT : ARRAY[1..6] OF ST_RCON_Direct_OUT_Axis;  (* RCON1 6軸分 PLC→RCON 指令（内部変数・通信変換は別途） *)
    RCON1_PowerStateRaw : ARRAY[0..4] OF WORD;  (* RCON1：入力IN02～06の正規化済み生ワード。詳細意味は構成依存。 *)
    RCON1_RxRaw : ARRAY[0..71] OF UINT;  (* RCON1：E001入力を読取った通信値。書換えない。 *)
    RCON1_RxWord : ARRAY[0..71] OF WORD;  (* RCON1：バイト順を正規化した論理入力ワード。 *)
    RCON1_SpeedUnit_mm_s : LREAL;  (* RCON1 速度の1カウント量mm/s。実機設定1.0または0.1を確認。未確認・0では使用しない。 *)
    RCON1_SwapBytes : BOOL;  (* RCON1：初期FALSEは仮値。1ワード内のバイト交換が必要か実機で確認。 *)
    RCON1_TxUInt : ARRAY[0..55] OF UINT;  (* RCON1：バイト順を適用した送信候補。実I/Oそのものではない。 *)
    RCON1_TxWord : ARRAY[0..55] OF WORD;  (* RCON1：内部値から作成した論理出力ワード。 *)
    RCON1_WriteEnable : BOOL;  (* RCON1：初期FALSE。実出力への書込みを許可。OFFは出力更新保留であり停止ではない。 *)
    RCON2_AxisApply : ARRAY[1..5] OF BOOL;  (* RCON2：初期FALSE。指定軸の8ワードを書込む。OFFは停止ではない。 *)
    RCON2_AxisLinked : ARRAY[1..5] OF BOOL;  (* RCON2：入力：軸No.0～4のリンク状態。 *)
    RCON2_AxisWritten : ARRAY[1..5] OF BOOL;  (* RCON2：各軸出力へ代入したサイクルのみTRUE。RCON受付・完了ではない。 *)
    RCON2_ByteOrderConfirmed : BOOL;  (* RCON2：初期FALSE。既知の位置とbitでワード順・バイト順を確認して設定。 *)
    RCON2_CommOK : BOOL;  (* RCON2：初期FALSE。CPUの実EtherCAT通信状態から別途作成。TRUE固定禁止。 *)
    RCON2_EncodeError : ARRAY[1..5] OF UINT;  (* RCON2：変換エラー番号。0正常、1単位、2位置、3幅、4速度、5加減速、6押付け、7両方向ジョグ。 *)
    RCON2_EncodeOK : ARRAY[1..5] OF BOOL;  (* RCON2：通信形式へ数値変換できたか。安全・運転許可ではない。 *)
    RCON2_GwAlarmCode : UINT;  (* RCON2：入力：ゲートウェイALMCの下位8bit。軸AlarmCodeとは別。 *)
    RCON2_GwApply : BOOL;  (* RCON2：初期FALSE。共通MON/RTEワードを書込む。 *)
    RCON2_GwAxisCommError : BOOL;  (* RCON2：入力：ゲートウェイと軸の通信異常ERRT。 *)
    RCON2_GwControllerCommLatch : BOOL;  (* RCON2：入力：運転中ERR-C保持LERC。 *)
    RCON2_GwHeavyAlarm : BOOL;  (* RCON2：入力：再起動が必要なゲートウェイ異常ALMH。 *)
    RCON2_GwLightAlarm : BOOL;  (* RCON2：入力：ゲートウェイ軽微異常ALML。 *)
    RCON2_GwMON_Request : BOOL;  (* RCON2：初期FALSE。ゲートウェイMON要求。論理b15。安全停止ではない。 *)
    RCON2_GwManual : BOOL;  (* RCON2：入力：MANUスイッチ選択MOD。 *)
    RCON2_GwRTE_Request : BOOL;  (* RCON2：初期FALSE。ゲートウェイ通信異常ラッチ解除要求。論理b13。 *)
    RCON2_GwRun : BOOL;  (* RCON2：入力：ゲートウェイ正常動作中RUN。 *)
    RCON2_GwSystemStop : BOOL;  (* RCON2：入力：システムSTOP入力による停止状態SEMG。安全回路の代用不可。 *)
    RCON2_GwWritten : BOOL;  (* RCON2：共通出力へ代入したサイクルのみTRUE。RCON受付の意味ではない。 *)
    RCON2_IN : ARRAY[1..5] OF ST_RCON_Direct_IN_Axis;  (* RCON2 5軸分 RCON→PLC 取得値・状態（内部変数・通信変換は別途） *)
    RCON2_LayoutConfirmed : BOOL;  (* RCON2：初期FALSE。全5軸直接数値指定・共通8W・軸順・占有を確認して設定。 *)
    RCON2_MotionPermit : ARRAY[1..5] OF BOOL;  (* RCON2：初期FALSE。機械範囲・安全・運転条件から別途作成する運転許可。単純TRUE固定禁止。 *)
    RCON2_OUT : ARRAY[1..5] OF ST_RCON_Direct_OUT_Axis;  (* RCON2 5軸分 PLC→RCON 指令（内部変数・通信変換は別途） *)
    RCON2_PowerStateRaw : ARRAY[0..4] OF WORD;  (* RCON2：入力IN02～06の正規化済み生ワード。詳細意味は構成依存。 *)
    RCON2_RxRaw : ARRAY[0..47] OF UINT;  (* RCON2：E005（末尾_1）入力を読取った通信値。書換えない。 *)
    RCON2_RxWord : ARRAY[0..47] OF WORD;  (* RCON2：バイト順を正規化した論理入力ワード。 *)
    RCON2_SpeedUnit_mm_s : LREAL;  (* RCON2 速度の1カウント量mm/s。実機設定1.0または0.1を確認。未確認・0では使用しない。 *)
    RCON2_SwapBytes : BOOL;  (* RCON2：初期FALSEは仮値。1ワード内のバイト交換が必要か実機で確認。 *)
    RCON2_TxUInt : ARRAY[0..47] OF UINT;  (* RCON2：バイト順を適用した送信候補。実I/Oそのものではない。 *)
    RCON2_TxWord : ARRAY[0..47] OF WORD;  (* RCON2：内部値から作成した論理出力ワード。 *)
    RCON2_WriteEnable : BOOL;  (* RCON2：初期FALSE。実出力への書込みを許可。OFFは出力更新保留であり停止ではない。 *)
END_VAR
VAR
    _e1 : R_TRIG;
    _p2 : BOOL;
    _e3 : R_TRIG;
    _p4 : BOOL;
    _e5 : R_TRIG;
    _p6 : BOOL;
    _e7 : R_TRIG;
    _e8 : R_TRIG;
    _p9 : BOOL;
    _e10 : R_TRIG;
    _e11 : R_TRIG;
    _p12 : BOOL;
    _p13 : BOOL;
END_VAR

(* Section RCON_IAI: ladder, written here as Structured Text *)

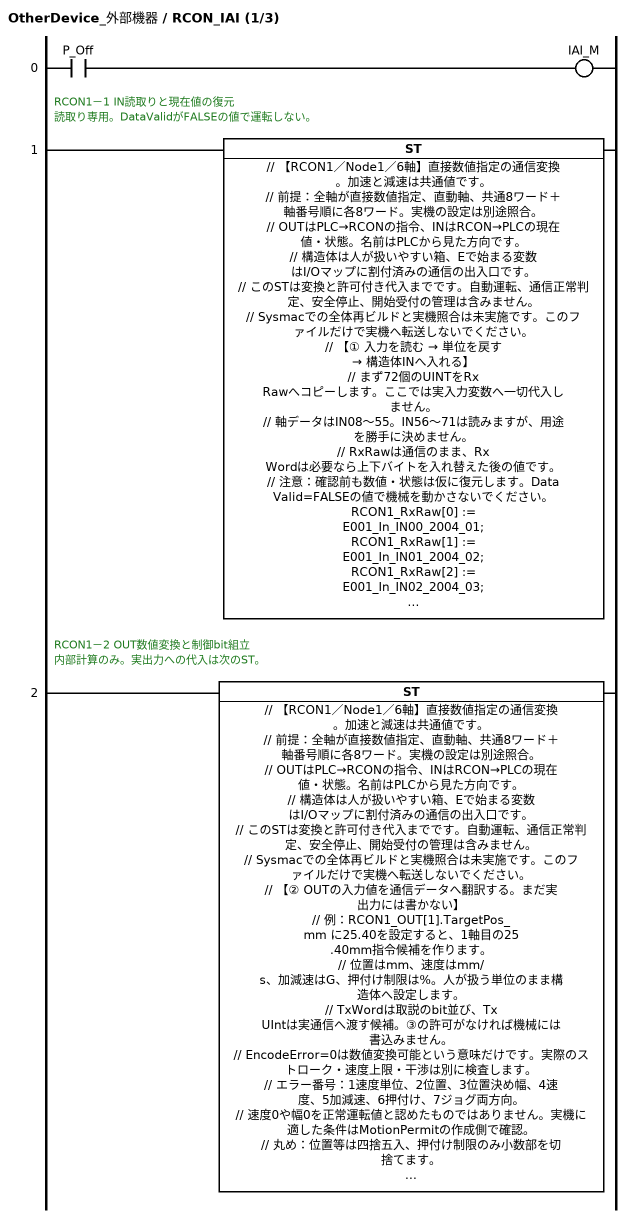
(* Rung 0 *)
IAI_M := P_Off;
(* Rung 1: RCON1－1 IN読取りと現在値の復元 / 読取り専用。DataValidがFALSEの値で運転しない。 *)
// 【RCON1／Node1／6軸】直接数値指定の通信変換。加速と減速は共通値です。
// 前提：全軸が直接数値指定、直動軸、共通8ワード＋軸番号順に各8ワード。実機の設定は別途照合。
// OUTはPLC→RCONの指令、INはRCON→PLCの現在値・状態。名前はPLCから見た方向です。
// 構造体は人が扱いやすい箱、Eで始まる変数はI/Oマップに割付済みの通信の出入口です。
// このSTは変換と許可付き代入までです。自動運転、通信正常判定、安全停止、開始受付の管理は含みません。
// Sysmacでの全体再ビルドと実機照合は未実施です。このファイルだけで実機へ転送しないでください。
// 【① 入力を読む → 単位を戻す → 構造体INへ入れる】
// まず72個のUINTをRxRawへコピーします。ここでは実入力変数へ一切代入しません。
// 軸データはIN08～55。IN56～71は読みますが、用途を勝手に決めません。
// RxRawは通信のまま、RxWordは必要なら上下バイトを入れ替えた後の値です。
// 注意：確認前も数値・状態は仮に復元します。DataValid=FALSEの値で機械を動かさないでください。
RCON1_RxRaw[0] := E001_In_IN00_2004_01;
RCON1_RxRaw[1] := E001_In_IN01_2004_02;
RCON1_RxRaw[2] := E001_In_IN02_2004_03;
RCON1_RxRaw[3] := E001_In_IN03_2004_04;
RCON1_RxRaw[4] := E001_In_IN04_2004_05;
RCON1_RxRaw[5] := E001_In_IN05_2004_06;
RCON1_RxRaw[6] := E001_In_IN06_2004_07;
RCON1_RxRaw[7] := E001_In_IN07_2004_08;
RCON1_RxRaw[8] := E001_In_IN08_2004_09;
RCON1_RxRaw[9] := E001_In_IN09_2004_0A;
RCON1_RxRaw[10] := E001_In_IN10_2004_0B;
RCON1_RxRaw[11] := E001_In_IN11_2004_0C;
RCON1_RxRaw[12] := E001_In_IN12_2004_0D;
RCON1_RxRaw[13] := E001_In_IN13_2004_0E;
RCON1_RxRaw[14] := E001_In_IN14_2004_0F;
RCON1_RxRaw[15] := E001_In_IN15_2004_10;
RCON1_RxRaw[16] := E001_In_IN16_2004_11;
RCON1_RxRaw[17] := E001_In_IN17_2004_12;
RCON1_RxRaw[18] := E001_In_IN18_2004_13;
RCON1_RxRaw[19] := E001_In_IN19_2004_14;
RCON1_RxRaw[20] := E001_In_IN20_2004_15;
RCON1_RxRaw[21] := E001_In_IN21_2004_16;
RCON1_RxRaw[22] := E001_In_IN22_2004_17;
RCON1_RxRaw[23] := E001_In_IN23_2004_18;
RCON1_RxRaw[24] := E001_In_IN24_2004_19;
RCON1_RxRaw[25] := E001_In_IN25_2004_1A;
RCON1_RxRaw[26] := E001_In_IN26_2004_1B;
RCON1_RxRaw[27] := E001_In_IN27_2004_1C;
RCON1_RxRaw[28] := E001_In_IN28_2004_1D;
RCON1_RxRaw[29] := E001_In_IN29_2004_1E;
RCON1_RxRaw[30] := E001_In_IN30_2004_1F;
RCON1_RxRaw[31] := E001_In_IN31_2004_20;
RCON1_RxRaw[32] := E001_In_IN32_2004_21;
RCON1_RxRaw[33] := E001_In_IN33_2004_22;
RCON1_RxRaw[34] := E001_In_IN34_2004_23;
RCON1_RxRaw[35] := E001_In_IN35_2004_24;
RCON1_RxRaw[36] := E001_In_IN36_2004_25;
RCON1_RxRaw[37] := E001_In_IN37_2004_26;
RCON1_RxRaw[38] := E001_In_IN38_2004_27;
RCON1_RxRaw[39] := E001_In_IN39_2004_28;
RCON1_RxRaw[40] := E001_In_IN40_2004_29;
RCON1_RxRaw[41] := E001_In_IN41_2004_2A;
RCON1_RxRaw[42] := E001_In_IN42_2004_2B;
RCON1_RxRaw[43] := E001_In_IN43_2004_2C;
RCON1_RxRaw[44] := E001_In_IN44_2004_2D;
RCON1_RxRaw[45] := E001_In_IN45_2004_2E;
RCON1_RxRaw[46] := E001_In_IN46_2004_2F;
RCON1_RxRaw[47] := E001_In_IN47_2004_30;
RCON1_RxRaw[48] := E001_In_IN48_2004_31;
RCON1_RxRaw[49] := E001_In_IN49_2004_32;
RCON1_RxRaw[50] := E001_In_IN50_2004_33;
RCON1_RxRaw[51] := E001_In_IN51_2004_34;
RCON1_RxRaw[52] := E001_In_IN52_2004_35;
RCON1_RxRaw[53] := E001_In_IN53_2004_36;
RCON1_RxRaw[54] := E001_In_IN54_2004_37;
RCON1_RxRaw[55] := E001_In_IN55_2004_38;
RCON1_RxRaw[56] := E001_In_IN56_2004_39;
RCON1_RxRaw[57] := E001_In_IN57_2004_3A;
RCON1_RxRaw[58] := E001_In_IN58_2004_3B;
RCON1_RxRaw[59] := E001_In_IN59_2004_3C;
RCON1_RxRaw[60] := E001_In_IN60_2004_3D;
RCON1_RxRaw[61] := E001_In_IN61_2004_3E;
RCON1_RxRaw[62] := E001_In_IN62_2004_3F;
RCON1_RxRaw[63] := E001_In_IN63_2004_40;
RCON1_RxRaw[64] := E001_In_IN64_2004_41;
RCON1_RxRaw[65] := E001_In_IN65_2004_42;
RCON1_RxRaw[66] := E001_In_IN66_2004_43;
RCON1_RxRaw[67] := E001_In_IN67_2004_44;
RCON1_RxRaw[68] := E001_In_IN68_2004_45;
RCON1_RxRaw[69] := E001_In_IN69_2004_46;
RCON1_RxRaw[70] := E001_In_IN70_2004_47;
RCON1_RxRaw[71] := E001_In_IN71_2004_48;

// 取説の論理ワードへ正規化。Swapは1ワード内の上下バイト交換です。
// SwapBytesは推測で設定せず、既知の位置とbitで実機照合してください。
FOR ConvWordIndex := INT#0 TO INT#71 DO
    RCON1_RxWord[ConvWordIndex] := UINT_TO_WORD(RCON1_RxRaw[ConvWordIndex]);
    IF RCON1_SwapBytes THEN
        RCON1_RxWord[ConvWordIndex] := Swap(RCON1_RxWord[ConvWordIndex]);
    END_IF;
END_FOR;

ConvUnitOK := (RCON1_SpeedUnit_mm_s = LREAL#1.0) OR
              (RCON1_SpeedUnit_mm_s = LREAL#0.1);

// 【①-2 共通状態】IN00はユニット全体、IN01は各軸のリンク情報です。
// TestABit(ワード, bit番号)は、そのスイッチがONかをBOOLで取り出す命令です。
// 例：IN01のb0は軸No.0→配列[1]、b1は軸No.1→配列[2]。配列番号と実機軸番号は1違います。
// 共通固定領域。ここで使うbit番号は取説の論理bitです（MJ0384 6-24～6-25）。
RCON1_GwRun := TestABit(RCON1_RxWord[0], USINT#15);
RCON1_GwControllerCommLatch := TestABit(RCON1_RxWord[0], USINT#14);
RCON1_GwAxisCommError := TestABit(RCON1_RxWord[0], USINT#13);
RCON1_GwManual := TestABit(RCON1_RxWord[0], USINT#12);
RCON1_GwHeavyAlarm := TestABit(RCON1_RxWord[0], USINT#11);
RCON1_GwLightAlarm := TestABit(RCON1_RxWord[0], USINT#10);
RCON1_GwSystemStop := TestABit(RCON1_RxWord[0], USINT#8);
RCON1_GwAlarmCode := WORD_TO_UINT(RCON1_RxWord[0] AND WORD#16#00FF);
FOR ConvWordIndex := INT#0 TO INT#4 DO
    RCON1_PowerStateRaw[ConvWordIndex] := RCON1_RxWord[ConvWordIndex + INT#2];
END_FOR;

// 【①-3 軸ごとに同じ読取りを繰り返す】
// FORは1～6軸を順番に処理します。ConvBaseはその軸の先頭番号です。
// 計算：8+(軸番号-1)×8。1軸目=8、2軸目=16、3軸目=24。先頭8ワードは共通領域です。
FOR ConvAxisIndex := INT#1 TO INT#6 DO
    ConvBase := INT#8 + (ConvAxisIndex - INT#1) * INT#8;
    RCON1_AxisLinked[ConvAxisIndex] :=
        TestABit(RCON1_RxWord[1], INT_TO_USINT(ConvAxisIndex - INT#1));

// 例：下位2540／上位0なら32bit値2540→25.40mm。
// 上位を16bit左に動かして下位とORで重ねます。SHLが左シフト、ORがビットの合成です。
// 負位置はDWORD_TO_DINTで符号を復元。下位62996／上位65535なら-2540→-25.40mm。
    // 現在位置：下位・上位を結合、符号付き32bitとして解釈、0.01mmをmmへ。
    ConvDWord := SHL(WORD_TO_DWORD(RCON1_RxWord[ConvBase + INT#1]), ULINT#16)
                 OR WORD_TO_DWORD(RCON1_RxWord[ConvBase]);
    RCON1_IN[ConvAxisIndex].ActualPos_mm :=
        DINT_TO_LREAL(DWORD_TO_DINT(ConvDWord)) * LREAL#0.01;

    // 電流：32bitのmA。RCON-PCでは指令電流であり、実測トルクではありません。
    ConvDWord := SHL(WORD_TO_DWORD(RCON1_RxWord[ConvBase + INT#3]), ULINT#16)
                 OR WORD_TO_DWORD(RCON1_RxWord[ConvBase + INT#2]);
    RCON1_IN[ConvAxisIndex].Current_mA := DWORD_TO_DINT(ConvDWord);

    // 現在速度：16bitの負数をINTとして読む。UINTのまま速度にしません。
    IF ConvUnitOK THEN
        RCON1_IN[ConvAxisIndex].ActualSpeed_mm_s :=
            INT_TO_LREAL(WORD_TO_INT(RCON1_RxWord[ConvBase + INT#4])) * RCON1_SpeedUnit_mm_s;
    END_IF;
    // 単位不明のとき速度は前値を保持し、DataValidはFALSEにします。
    // 軸内の+5ワードは予約のため値を使用しません。
    RCON1_IN[ConvAxisIndex].AlarmCode := WORD_TO_UINT(RCON1_RxWord[ConvBase + INT#6]);

// 例：Status.ServoReady=TRUEは「サーボON状態を受信した」という意味。
// OUT側Control.ServoOn=TRUEは「サーボONを要求する」という意味で、指令と結果を区別します。
    // 状態ワード：12個のBOOLへ分解。予約b6,b9～11は使いません。
    RCON1_IN[ConvAxisIndex].Status.PositionDone := TestABit(RCON1_RxWord[ConvBase + INT#7], USINT#0);
    RCON1_IN[ConvAxisIndex].Status.HomeDone := TestABit(RCON1_RxWord[ConvBase + INT#7], USINT#1);
    RCON1_IN[ConvAxisIndex].Status.Moving := TestABit(RCON1_RxWord[ConvBase + INT#7], USINT#2);
    RCON1_IN[ConvAxisIndex].Status.Alarm := TestABit(RCON1_RxWord[ConvBase + INT#7], USINT#3);
    RCON1_IN[ConvAxisIndex].Status.ServoReady := TestABit(RCON1_RxWord[ConvBase + INT#7], USINT#4);
    RCON1_IN[ConvAxisIndex].Status.PushMiss := TestABit(RCON1_RxWord[ConvBase + INT#7], USINT#5);
    RCON1_IN[ConvAxisIndex].Status.OverloadWarning := TestABit(RCON1_RxWord[ConvBase + INT#7], USINT#7);
    RCON1_IN[ConvAxisIndex].Status.CommandDone := TestABit(RCON1_RxWord[ConvBase + INT#7], USINT#8);
    RCON1_IN[ConvAxisIndex].Status.Zone1 := TestABit(RCON1_RxWord[ConvBase + INT#7], USINT#12);
    RCON1_IN[ConvAxisIndex].Status.Zone2 := TestABit(RCON1_RxWord[ConvBase + INT#7], USINT#13);
    RCON1_IN[ConvAxisIndex].Status.ControllerReady := TestABit(RCON1_RxWord[ConvBase + INT#7], USINT#14);
    RCON1_IN[ConvAxisIndex].Status.EmergencyStop := TestABit(RCON1_RxWord[ConvBase + INT#7], USINT#15);

    // DataValidは直接受信bitではなく、今回の内部設計で決めた内部判定です。
    // CommOKはCPUの実通信状態から別途作成。単にTRUE固定にしないでください。
    // DataValidは運転許可や安全保証ではありません。各異常・原点等は別途確認。
    RCON1_IN[ConvAxisIndex].DataValid := RCON1_CommOK AND RCON1_LayoutConfirmed
        AND RCON1_ByteOrderConfirmed AND ConvUnitOK AND RCON1_GwRun
        AND RCON1_AxisLinked[ConvAxisIndex] AND NOT RCON1_GwAxisCommError;
END_FOR;
(* Rung 2: RCON1－2 OUT数値変換と制御bit組立 / 内部計算のみ。実出力への代入は次のST。 *)
// 【RCON1／Node1／6軸】直接数値指定の通信変換。加速と減速は共通値です。
// 前提：全軸が直接数値指定、直動軸、共通8ワード＋軸番号順に各8ワード。実機の設定は別途照合。
// OUTはPLC→RCONの指令、INはRCON→PLCの現在値・状態。名前はPLCから見た方向です。
// 構造体は人が扱いやすい箱、Eで始まる変数はI/Oマップに割付済みの通信の出入口です。
// このSTは変換と許可付き代入までです。自動運転、通信正常判定、安全停止、開始受付の管理は含みません。
// Sysmacでの全体再ビルドと実機照合は未実施です。このファイルだけで実機へ転送しないでください。
// 【② OUTの入力値を通信データへ翻訳する。まだ実出力には書かない】
// 例：RCON1_OUT[1].TargetPos_mm に25.40を設定すると、1軸目の25.40mm指令候補を作ります。
// 位置はmm、速度はmm/s、加減速はG、押付け制限は%。人が扱う単位のまま構造体へ設定します。
// TxWordは取説のbit並び、TxUIntは実通信へ渡す候補。③の許可がなければ機械には書込みません。
// EncodeError=0は数値変換可能という意味だけです。実際のストローク・速度上限・干渉は別に検査します。
// エラー番号：1速度単位、2位置、3位置決め幅、4速度、5加減速、6押付け、7ジョグ両方向。
// 速度0や幅0を正常運転値と認めたものではありません。実機に適した条件はMotionPermitの作成側で確認。
// 丸め：位置等は四捨五入、押付け制限のみ小数部を切捨てます。

ConvUnitOK := (RCON1_SpeedUnit_mm_s = LREAL#1.0) OR
              (RCON1_SpeedUnit_mm_s = LREAL#0.1);

// 共通制御：MONは論理b15、RTEは論理b13。他のbitは0。
// MONを落とす処理を安全停止として扱わないでください。
RCON1_TxWord[0] := WORD#16#0000;
IF RCON1_GwMON_Request THEN
    RCON1_TxWord[0] := RCON1_TxWord[0] OR WORD#16#8000;
END_IF;
IF RCON1_GwRTE_Request THEN
    RCON1_TxWord[0] := RCON1_TxWord[0] OR WORD#16#2000;
END_IF;

FOR ConvAxisIndex := INT#1 TO INT#6 DO
    ConvBase := INT#8 + (ConvAxisIndex - INT#1) * INT#8;
    RCON1_EncodeError[ConvAxisIndex] := UINT#0;

    // 比較で範囲を確認してから型変換するため、NaN・無限大も変換対象から外れます。
    // 位置・幅9999.99mmはこの案で採用する通信範囲の上限で、実機ストロークではありません。
    IF NOT ConvUnitOK THEN
        RCON1_EncodeError[ConvAxisIndex] := UINT#1;
    ELSIF NOT ((RCON1_OUT[ConvAxisIndex].TargetPos_mm >= LREAL#-9999.99) AND
               (RCON1_OUT[ConvAxisIndex].TargetPos_mm <= LREAL#9999.99)) THEN
        RCON1_EncodeError[ConvAxisIndex] := UINT#2;
    ELSIF NOT ((RCON1_OUT[ConvAxisIndex].PositionBand_mm >= LREAL#0.0) AND
               (RCON1_OUT[ConvAxisIndex].PositionBand_mm <= LREAL#9999.99)) THEN
        RCON1_EncodeError[ConvAxisIndex] := UINT#3;
    ELSIF NOT ((RCON1_OUT[ConvAxisIndex].Speed_mm_s >= LREAL#0.0) AND
               (RCON1_OUT[ConvAxisIndex].Speed_mm_s <= LREAL#65535.0 * RCON1_SpeedUnit_mm_s)) THEN
        RCON1_EncodeError[ConvAxisIndex] := UINT#4;
    ELSIF NOT ((RCON1_OUT[ConvAxisIndex].AccDec_G >= LREAL#0.0) AND
               (RCON1_OUT[ConvAxisIndex].AccDec_G <= LREAL#655.35)) THEN
        RCON1_EncodeError[ConvAxisIndex] := UINT#5;
    ELSIF NOT ((RCON1_OUT[ConvAxisIndex].PushLimit_pct >= LREAL#0.0) AND
               (RCON1_OUT[ConvAxisIndex].PushLimit_pct <= LREAL#200.0)) THEN
        RCON1_EncodeError[ConvAxisIndex] := UINT#6;
    ELSIF RCON1_OUT[ConvAxisIndex].Control.JogMinus AND RCON1_OUT[ConvAxisIndex].Control.JogPlus THEN
        RCON1_EncodeError[ConvAxisIndex] := UINT#7;
    END_IF;

    RCON1_EncodeOK[ConvAxisIndex] := RCON1_EncodeError[ConvAxisIndex] = UINT#0;
    IF RCON1_EncodeOK[ConvAxisIndex] THEN
    // 【数値例】TargetPos_mm=25.40→×100で2540。下位ワード2540、上位ワード0。
// 700.25mm→70025なので下位4489、上位1。65536を超えた分が上位に入ります。
// DINTは符号付きの数、DWORDは同じ32bitの模様。負数の符号を壊さず分割するために使い分けます。
// TRUNCは小数部を捨てます。正数+0.5／負数-0.5を先に行い、四捨五入を明示しています。
    // 目標位置：mmから0.01mmの符号付き整数へ。
        ConvScaled := RCON1_OUT[ConvAxisIndex].TargetPos_mm * LREAL#100.0;
        IF ConvScaled >= LREAL#0.0 THEN
            ConvPos := LINT_TO_DINT(TRUNC(ConvScaled + LREAL#0.5));
        ELSE
            ConvPos := LINT_TO_DINT(TRUNC(ConvScaled - LREAL#0.5));
        END_IF;
        // 負数を含む32bitパターンを保ち、下位・上位の16bitへ分割。
        ConvDWord := DINT_TO_DWORD(ConvPos);
        RCON1_TxWord[ConvBase] := DWORD_TO_WORD(ConvDWord AND DWORD#16#0000FFFF);
        RCON1_TxWord[ConvBase + INT#1] := DWORD_TO_WORD(SHR(ConvDWord, ULINT#16));

        // 位置決め幅：非負の内部整数としてUDINTを選定（メーカーの符号なし保証ではありません）。
        ConvBand := LINT_TO_UDINT(TRUNC(RCON1_OUT[ConvAxisIndex].PositionBand_mm * LREAL#100.0 + LREAL#0.5));
        ConvDWord := UDINT_TO_DWORD(ConvBand);
        RCON1_TxWord[ConvBase + INT#2] := DWORD_TO_WORD(ConvDWord AND DWORD#16#0000FFFF);
        RCON1_TxWord[ConvBase + INT#3] := DWORD_TO_WORD(SHR(ConvDWord, ULINT#16));

// 速度20mm/s：速度単位1.0なら20、0.1なら200を送信します。
// 加減速0.20G：×100して20。加速と減速の両方に同じ値を使います。
// 押付け50%：×255÷100=127.5を切捨てて127。押付けの使用可否・上限は実機仕様で別確認。
        // 速度は1カウント量が1.0か0.1かで値が10倍変わります。
        ConvSpeed := LINT_TO_UINT(TRUNC(RCON1_OUT[ConvAxisIndex].Speed_mm_s / RCON1_SpeedUnit_mm_s + LREAL#0.5));
        ConvAccDec := LINT_TO_UINT(TRUNC(RCON1_OUT[ConvAxisIndex].AccDec_G * LREAL#100.0 + LREAL#0.5));
        ConvPush := LINT_TO_UINT(TRUNC(RCON1_OUT[ConvAxisIndex].PushLimit_pct * LREAL#255.0 / LREAL#100.0));
        RCON1_TxWord[ConvBase + INT#4] := UINT_TO_WORD(ConvSpeed);
        RCON1_TxWord[ConvBase + INT#5] := UINT_TO_WORD(ConvAccDec);
        RCON1_TxWord[ConvBase + INT#6] := UINT_TO_WORD(ConvPush);
    END_IF;
    // 不正値の場合、数値ワードは前値保持。EncodeOK=FALSEで03の書込みを抑止。
    // 前値保持は停止指令ではありません。停止・異常処理は別途設計してください。

    // Controlを論理bitへ詰める。予約b9は必ず0。
    RCON1_TxWord[ConvBase + INT#7] := WORD#16#0000;
// b0 DSTR／Control.Start：TRUEで開始要求。受付応答と10ms以上の保持を確認してOFF。常時ONにしない。
    IF RCON1_OUT[ConvAxisIndex].Control.Start THEN
        RCON1_TxWord[ConvBase + INT#7] := RCON1_TxWord[ConvBase + INT#7] OR WORD#16#0001;
    END_IF;
// b1 HOME／Control.Home：TRUEで原点復帰を指令。原点復帰完了はIN側HomeDoneで確認。
    IF RCON1_OUT[ConvAxisIndex].Control.Home THEN
        RCON1_TxWord[ConvBase + INT#7] := RCON1_TxWord[ConvBase + INT#7] OR WORD#16#0002;
    END_IF;
// b2 STP／Control.Pause：TRUEで一時停止、FALSEで解除。非常停止・安全停止の代用ではない。
    IF RCON1_OUT[ConvAxisIndex].Control.Pause THEN
        RCON1_TxWord[ConvBase + INT#7] := RCON1_TxWord[ConvBase + INT#7] OR WORD#16#0004;
    END_IF;
// b3 RES／Control.Reset：TRUEでアラームリセット要求。コールドスタート級の異常には使用できない。
    IF RCON1_OUT[ConvAxisIndex].Control.Reset THEN
        RCON1_TxWord[ConvBase + INT#7] := RCON1_TxWord[ConvBase + INT#7] OR WORD#16#0008;
    END_IF;
// b4 SON／Control.ServoOn：TRUEでサーボON要求。ON状態はIN側ServoReadyで確認。
    IF RCON1_OUT[ConvAxisIndex].Control.ServoOn THEN
        RCON1_TxWord[ConvBase + INT#7] := RCON1_TxWord[ConvBase + INT#7] OR WORD#16#0010;
    END_IF;
// b5 JISL／Control.InchingSelect：TRUEは一定距離のインチング、FALSEは押している間のジョグ。
    IF RCON1_OUT[ConvAxisIndex].Control.InchingSelect THEN
        RCON1_TxWord[ConvBase + INT#7] := RCON1_TxWord[ConvBase + INT#7] OR WORD#16#0020;
    END_IF;
// b6 JVEL／Control.JogSpeedSelect：FALSEは速度No.26・距離No.48、TRUEは速度No.47または指令速度・距離No.49。
    IF RCON1_OUT[ConvAxisIndex].Control.JogSpeedSelect THEN
        RCON1_TxWord[ConvBase + INT#7] := RCON1_TxWord[ConvBase + INT#7] OR WORD#16#0040;
    END_IF;
// b7 JOG-／Control.JogMinus：TRUEで原点方向へジョグ。反対方向指令との同時ONを防ぐ。
    IF RCON1_OUT[ConvAxisIndex].Control.JogMinus THEN
        RCON1_TxWord[ConvBase + INT#7] := RCON1_TxWord[ConvBase + INT#7] OR WORD#16#0080;
    END_IF;
// b8 JOG+／Control.JogPlus：TRUEで反原点方向へジョグ。反対方向指令との同時ONを防ぐ。
    IF RCON1_OUT[ConvAxisIndex].Control.JogPlus THEN
        RCON1_TxWord[ConvBase + INT#7] := RCON1_TxWord[ConvBase + INT#7] OR WORD#16#0100;
    END_IF;
// b10 GSL0／Control.GainSelect0：GainSelect1と組合せてサーボゲインセット0～3を選ぶ。機械調整用。
    IF RCON1_OUT[ConvAxisIndex].Control.GainSelect0 THEN
        RCON1_TxWord[ConvBase + INT#7] := RCON1_TxWord[ConvBase + INT#7] OR WORD#16#0400;
    END_IF;
// b11 GSL1／Control.GainSelect1：GainSelect0との2bitで選択。速度指令とは別の機能。
    IF RCON1_OUT[ConvAxisIndex].Control.GainSelect1 THEN
        RCON1_TxWord[ConvBase + INT#7] := RCON1_TxWord[ConvBase + INT#7] OR WORD#16#0800;
    END_IF;
// b12 PUSH／Control.PushEnable：TRUEは押付け、FALSEは通常位置決め。押付け条件は別途確認。
    IF RCON1_OUT[ConvAxisIndex].Control.PushEnable THEN
        RCON1_TxWord[ConvBase + INT#7] := RCON1_TxWord[ConvBase + INT#7] OR WORD#16#1000;
    END_IF;
// b13 DIR／Control.PushDirection：CON方式押付け時、TRUEは反原点方向、FALSEは原点方向。
    IF RCON1_OUT[ConvAxisIndex].Control.PushDirection THEN
        RCON1_TxWord[ConvBase + INT#7] := RCON1_TxWord[ConvBase + INT#7] OR WORD#16#2000;
    END_IF;
// b14 INC／Control.RelativeMove：FALSEは絶対座標、TRUEは現在位置からの相対移動量。
    IF RCON1_OUT[ConvAxisIndex].Control.RelativeMove THEN
        RCON1_TxWord[ConvBase + INT#7] := RCON1_TxWord[ConvBase + INT#7] OR WORD#16#4000;
    END_IF;
// b15 BKRL／Control.BrakeRelease：TRUEはブレーキ強制解除。通常FALSE。縦軸では落下等の危険がある。
    IF RCON1_OUT[ConvAxisIndex].Control.BrakeRelease THEN
        RCON1_TxWord[ConvBase + INT#7] := RCON1_TxWord[ConvBase + INT#7] OR WORD#16#8000;
    END_IF;
END_FOR;

// 論理ワードから実際に送るUINTへ。INと同じ1ワード内のバイト交換を適用します。
FOR ConvWordIndex := INT#0 TO INT#55 DO
    ConvWord := RCON1_TxWord[ConvWordIndex];
    IF RCON1_SwapBytes THEN
        ConvWord := Swap(ConvWord);
    END_IF;
    RCON1_TxUInt[ConvWordIndex] := WORD_TO_UINT(ConvWord);
END_FOR;

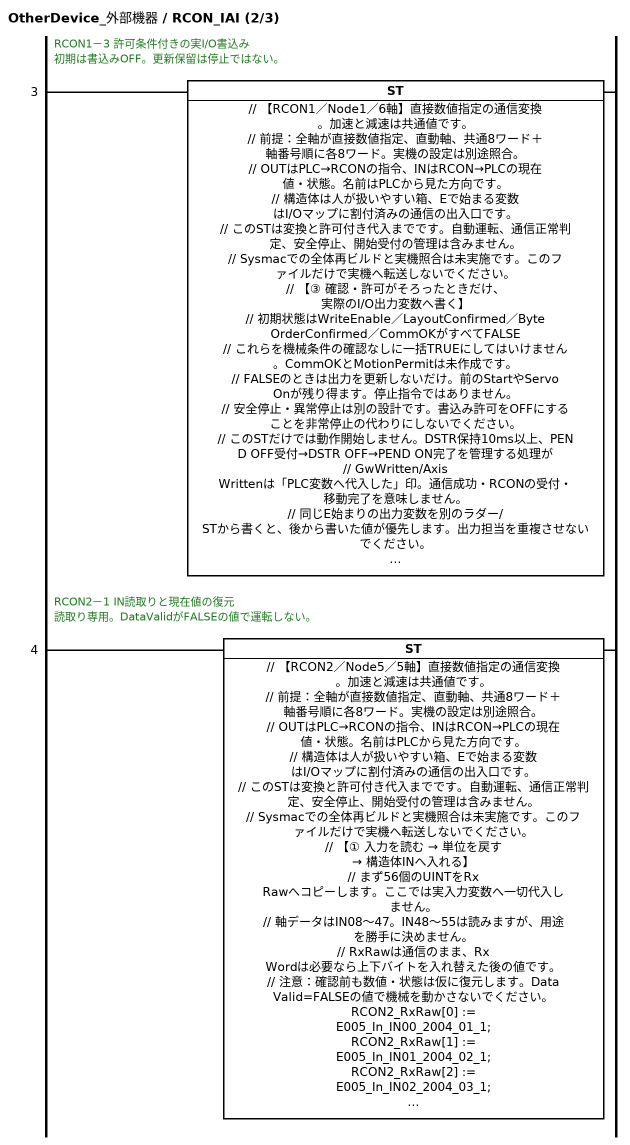
(* Rung 3: RCON1－3 許可条件付きの実I/O書込み / 初期は書込みOFF。更新保留は停止ではない。 *)
// 【RCON1／Node1／6軸】直接数値指定の通信変換。加速と減速は共通値です。
// 前提：全軸が直接数値指定、直動軸、共通8ワード＋軸番号順に各8ワード。実機の設定は別途照合。
// OUTはPLC→RCONの指令、INはRCON→PLCの現在値・状態。名前はPLCから見た方向です。
// 構造体は人が扱いやすい箱、Eで始まる変数はI/Oマップに割付済みの通信の出入口です。
// このSTは変換と許可付き代入までです。自動運転、通信正常判定、安全停止、開始受付の管理は含みません。
// Sysmacでの全体再ビルドと実機照合は未実施です。このファイルだけで実機へ転送しないでください。
// 【③ 確認・許可がそろったときだけ、実際のI/O出力変数へ書く】
// 初期状態はWriteEnable／LayoutConfirmed／ByteOrderConfirmed／CommOKがすべてFALSEです。
// これらを機械条件の確認なしに一括TRUEにしてはいけません。CommOKとMotionPermitは未作成です。
// FALSEのときは出力を更新しないだけ。前のStartやServoOnが残り得ます。停止指令ではありません。
// 安全停止・異常停止は別の設計です。書込み許可をOFFにすることを非常停止の代わりにしないでください。
// このSTだけでは動作開始しません。DSTR保持10ms以上、PEND OFF受付→DSTR OFF→PEND ON完了を管理する処理が必要です。
// GwWritten/AxisWrittenは「PLC変数へ代入した」印。通信成功・RCONの受付・移動完了を意味しません。
// 同じE始まりの出力変数を別のラダー/STから書くと、後から書いた値が優先します。出力担当を重複させないでください。

RCON1_GwWritten := FALSE;
FOR ConvAxisIndex := INT#1 TO INT#6 DO
    RCON1_AxisWritten[ConvAxisIndex] := FALSE;
END_FOR;

IF RCON1_WriteEnable AND RCON1_LayoutConfirmed AND RCON1_ByteOrderConfirmed AND RCON1_CommOK THEN
// 共通指令はMON/RTEのみ。最初のRUN応答に必要なため、軸DataValidとは別にGwApplyで許可します。
    IF RCON1_GwApply THEN
        E001_Out_OUT00_2003_01 := RCON1_TxUInt[0];
        RCON1_GwWritten := TRUE;
    END_IF;

// 1軸目＝実機軸No.0。OUT08～OUT15の8ワードをまとめて代入。
// AxisApply=この軸の更新許可、EncodeOK=変換OK、DataValid=入力情報の条件確認、MotionPermit=機械側の運転許可。
// 途中1ワードだけではなく、位置・幅・速度・加減速・押付け・制御を一組として渡します。
    IF RCON1_AxisApply[1] AND RCON1_EncodeOK[1] AND RCON1_IN[1].DataValid
       AND RCON1_MotionPermit[1] THEN
        E001_Out_OUT08_2003_09 := RCON1_TxUInt[8];
        E001_Out_OUT09_2003_0A := RCON1_TxUInt[9];
        E001_Out_OUT10_2003_0B := RCON1_TxUInt[10];
        E001_Out_OUT11_2003_0C := RCON1_TxUInt[11];
        E001_Out_OUT12_2003_0D := RCON1_TxUInt[12];
        E001_Out_OUT13_2003_0E := RCON1_TxUInt[13];
        E001_Out_OUT14_2003_0F := RCON1_TxUInt[14];
        E001_Out_OUT15_2003_10 := RCON1_TxUInt[15];
        RCON1_AxisWritten[1] := TRUE;
    END_IF;

// 2軸目＝実機軸No.1。OUT16～OUT23の8ワードをまとめて代入。
// AxisApply=この軸の更新許可、EncodeOK=変換OK、DataValid=入力情報の条件確認、MotionPermit=機械側の運転許可。
// 途中1ワードだけではなく、位置・幅・速度・加減速・押付け・制御を一組として渡します。
    IF RCON1_AxisApply[2] AND RCON1_EncodeOK[2] AND RCON1_IN[2].DataValid
       AND RCON1_MotionPermit[2] THEN
        E001_Out_OUT16_2003_11 := RCON1_TxUInt[16];
        E001_Out_OUT17_2003_12 := RCON1_TxUInt[17];
        E001_Out_OUT18_2003_13 := RCON1_TxUInt[18];
        E001_Out_OUT19_2003_14 := RCON1_TxUInt[19];
        E001_Out_OUT20_2003_15 := RCON1_TxUInt[20];
        E001_Out_OUT21_2003_16 := RCON1_TxUInt[21];
        E001_Out_OUT22_2003_17 := RCON1_TxUInt[22];
        E001_Out_OUT23_2003_18 := RCON1_TxUInt[23];
        RCON1_AxisWritten[2] := TRUE;
    END_IF;

// 3軸目＝実機軸No.2。OUT24～OUT31の8ワードをまとめて代入。
// AxisApply=この軸の更新許可、EncodeOK=変換OK、DataValid=入力情報の条件確認、MotionPermit=機械側の運転許可。
// 途中1ワードだけではなく、位置・幅・速度・加減速・押付け・制御を一組として渡します。
    IF RCON1_AxisApply[3] AND RCON1_EncodeOK[3] AND RCON1_IN[3].DataValid
       AND RCON1_MotionPermit[3] THEN
        E001_Out_OUT24_2003_19 := RCON1_TxUInt[24];
        E001_Out_OUT25_2003_1A := RCON1_TxUInt[25];
        E001_Out_OUT26_2003_1B := RCON1_TxUInt[26];
        E001_Out_OUT27_2003_1C := RCON1_TxUInt[27];
        E001_Out_OUT28_2003_1D := RCON1_TxUInt[28];
        E001_Out_OUT29_2003_1E := RCON1_TxUInt[29];
        E001_Out_OUT30_2003_1F := RCON1_TxUInt[30];
        E001_Out_OUT31_2003_20 := RCON1_TxUInt[31];
        RCON1_AxisWritten[3] := TRUE;
    END_IF;

// 4軸目＝実機軸No.3。OUT32～OUT39の8ワードをまとめて代入。
// AxisApply=この軸の更新許可、EncodeOK=変換OK、DataValid=入力情報の条件確認、MotionPermit=機械側の運転許可。
// 途中1ワードだけではなく、位置・幅・速度・加減速・押付け・制御を一組として渡します。
    IF RCON1_AxisApply[4] AND RCON1_EncodeOK[4] AND RCON1_IN[4].DataValid
       AND RCON1_MotionPermit[4] THEN
        E001_Out_OUT32_2003_21 := RCON1_TxUInt[32];
        E001_Out_OUT33_2003_22 := RCON1_TxUInt[33];
        E001_Out_OUT34_2003_23 := RCON1_TxUInt[34];
        E001_Out_OUT35_2003_24 := RCON1_TxUInt[35];
        E001_Out_OUT36_2003_25 := RCON1_TxUInt[36];
        E001_Out_OUT37_2003_26 := RCON1_TxUInt[37];
        E001_Out_OUT38_2003_27 := RCON1_TxUInt[38];
        E001_Out_OUT39_2003_28 := RCON1_TxUInt[39];
        RCON1_AxisWritten[4] := TRUE;
    END_IF;

// 5軸目＝実機軸No.4。OUT40～OUT47の8ワードをまとめて代入。
// AxisApply=この軸の更新許可、EncodeOK=変換OK、DataValid=入力情報の条件確認、MotionPermit=機械側の運転許可。
// 途中1ワードだけではなく、位置・幅・速度・加減速・押付け・制御を一組として渡します。
    IF RCON1_AxisApply[5] AND RCON1_EncodeOK[5] AND RCON1_IN[5].DataValid
       AND RCON1_MotionPermit[5] THEN
        E001_Out_OUT40_2003_29 := RCON1_TxUInt[40];
        E001_Out_OUT41_2003_2A := RCON1_TxUInt[41];
        E001_Out_OUT42_2003_2B := RCON1_TxUInt[42];
        E001_Out_OUT43_2003_2C := RCON1_TxUInt[43];
        E001_Out_OUT44_2003_2D := RCON1_TxUInt[44];
        E001_Out_OUT45_2003_2E := RCON1_TxUInt[45];
        E001_Out_OUT46_2003_2F := RCON1_TxUInt[46];
        E001_Out_OUT47_2003_30 := RCON1_TxUInt[47];
        RCON1_AxisWritten[5] := TRUE;
    END_IF;

// 6軸目＝実機軸No.5。OUT48～OUT55の8ワードをまとめて代入。
// AxisApply=この軸の更新許可、EncodeOK=変換OK、DataValid=入力情報の条件確認、MotionPermit=機械側の運転許可。
// 途中1ワードだけではなく、位置・幅・速度・加減速・押付け・制御を一組として渡します。
    IF RCON1_AxisApply[6] AND RCON1_EncodeOK[6] AND RCON1_IN[6].DataValid
       AND RCON1_MotionPermit[6] THEN
        E001_Out_OUT48_2003_31 := RCON1_TxUInt[48];
        E001_Out_OUT49_2003_32 := RCON1_TxUInt[49];
        E001_Out_OUT50_2003_33 := RCON1_TxUInt[50];
        E001_Out_OUT51_2003_34 := RCON1_TxUInt[51];
        E001_Out_OUT52_2003_35 := RCON1_TxUInt[52];
        E001_Out_OUT53_2003_36 := RCON1_TxUInt[53];
        E001_Out_OUT54_2003_37 := RCON1_TxUInt[54];
        E001_Out_OUT55_2003_38 := RCON1_TxUInt[55];
        RCON1_AxisWritten[6] := TRUE;
    END_IF;
END_IF;
// OUT01～07、OUT56～71は、このSTからは一切書き換えません。
// 現在の実機設定・別処理の用途が未確認なので、余剰領域を勝手にゼロクリアしません。
(* Rung 4: RCON2－1 IN読取りと現在値の復元 / 読取り専用。DataValidがFALSEの値で運転しない。 *)
// 【RCON2／Node5／5軸】直接数値指定の通信変換。加速と減速は共通値です。
// 前提：全軸が直接数値指定、直動軸、共通8ワード＋軸番号順に各8ワード。実機の設定は別途照合。
// OUTはPLC→RCONの指令、INはRCON→PLCの現在値・状態。名前はPLCから見た方向です。
// 構造体は人が扱いやすい箱、Eで始まる変数はI/Oマップに割付済みの通信の出入口です。
// このSTは変換と許可付き代入までです。自動運転、通信正常判定、安全停止、開始受付の管理は含みません。
// Sysmacでの全体再ビルドと実機照合は未実施です。このファイルだけで実機へ転送しないでください。
// 【① 入力を読む → 単位を戻す → 構造体INへ入れる】
// まず56個のUINTをRxRawへコピーします。ここでは実入力変数へ一切代入しません。
// 軸データはIN08～47。IN48～55は読みますが、用途を勝手に決めません。
// RxRawは通信のまま、RxWordは必要なら上下バイトを入れ替えた後の値です。
// 注意：確認前も数値・状態は仮に復元します。DataValid=FALSEの値で機械を動かさないでください。
RCON2_RxRaw[0] := E005_In_IN00_2004_01_1;
RCON2_RxRaw[1] := E005_In_IN01_2004_02_1;
RCON2_RxRaw[2] := E005_In_IN02_2004_03_1;
RCON2_RxRaw[3] := E005_In_IN03_2004_04_1;
RCON2_RxRaw[4] := E005_In_IN04_2004_05_1;
RCON2_RxRaw[5] := E005_In_IN05_2004_06_1;
RCON2_RxRaw[6] := E005_In_IN06_2004_07_1;
RCON2_RxRaw[7] := E005_In_IN07_2004_08_1;
RCON2_RxRaw[8] := E005_In_IN08_2004_09_1;
RCON2_RxRaw[9] := E005_In_IN09_2004_0A_1;
RCON2_RxRaw[10] := E005_In_IN10_2004_0B_1;
RCON2_RxRaw[11] := E005_In_IN11_2004_0C_1;
RCON2_RxRaw[12] := E005_In_IN12_2004_0D_1;
RCON2_RxRaw[13] := E005_In_IN13_2004_0E_1;
RCON2_RxRaw[14] := E005_In_IN14_2004_0F_1;
RCON2_RxRaw[15] := E005_In_IN15_2004_10_1;
RCON2_RxRaw[16] := E005_In_IN16_2004_11_1;
RCON2_RxRaw[17] := E005_In_IN17_2004_12_1;
RCON2_RxRaw[18] := E005_In_IN18_2004_13_1;
RCON2_RxRaw[19] := E005_In_IN19_2004_14_1;
RCON2_RxRaw[20] := E005_In_IN20_2004_15_1;
RCON2_RxRaw[21] := E005_In_IN21_2004_16_1;
RCON2_RxRaw[22] := E005_In_IN22_2004_17_1;
RCON2_RxRaw[23] := E005_In_IN23_2004_18_1;
RCON2_RxRaw[24] := E005_In_IN24_2004_19_1;
RCON2_RxRaw[25] := E005_In_IN25_2004_1A_1;
RCON2_RxRaw[26] := E005_In_IN26_2004_1B_1;
RCON2_RxRaw[27] := E005_In_IN27_2004_1C_1;
RCON2_RxRaw[28] := E005_In_IN28_2004_1D_1;
RCON2_RxRaw[29] := E005_In_IN29_2004_1E_1;
RCON2_RxRaw[30] := E005_In_IN30_2004_1F_1;
RCON2_RxRaw[31] := E005_In_IN31_2004_20_1;
RCON2_RxRaw[32] := E005_In_IN32_2004_21_1;
RCON2_RxRaw[33] := E005_In_IN33_2004_22_1;
RCON2_RxRaw[34] := E005_In_IN34_2004_23_1;
RCON2_RxRaw[35] := E005_In_IN35_2004_24_1;
RCON2_RxRaw[36] := E005_In_IN36_2004_25_1;
RCON2_RxRaw[37] := E005_In_IN37_2004_26_1;
RCON2_RxRaw[38] := E005_In_IN38_2004_27_1;
RCON2_RxRaw[39] := E005_In_IN39_2004_28_1;
RCON2_RxRaw[40] := E005_In_IN40_2004_29_1;
RCON2_RxRaw[41] := E005_In_IN41_2004_2A_1;
RCON2_RxRaw[42] := E005_In_IN42_2004_2B_1;
RCON2_RxRaw[43] := E005_In_IN43_2004_2C_1;
RCON2_RxRaw[44] := E005_In_IN44_2004_2D_1;
RCON2_RxRaw[45] := E005_In_IN45_2004_2E_1;
RCON2_RxRaw[46] := E005_In_IN46_2004_2F_1;
RCON2_RxRaw[47] := E005_In_IN47_2004_30_1;
RCON2_RxRaw[48] := E005_In_IN48_2004_31_1;
RCON2_RxRaw[49] := E005_In_IN49_2004_32_1;
RCON2_RxRaw[50] := E005_In_IN50_2004_33_1;
RCON2_RxRaw[51] := E005_In_IN51_2004_34_1;
RCON2_RxRaw[52] := E005_In_IN52_2004_35_1;
RCON2_RxRaw[53] := E005_In_IN53_2004_36_1;
RCON2_RxRaw[54] := E005_In_IN54_2004_37_1;
RCON2_RxRaw[55] := E005_In_IN55_2004_38_1;

// 取説の論理ワードへ正規化。Swapは1ワード内の上下バイト交換です。
// SwapBytesは推測で設定せず、既知の位置とbitで実機照合してください。
FOR ConvWordIndex := INT#0 TO INT#55 DO
    RCON2_RxWord[ConvWordIndex] := UINT_TO_WORD(RCON2_RxRaw[ConvWordIndex]);
    IF RCON2_SwapBytes THEN
        RCON2_RxWord[ConvWordIndex] := Swap(RCON2_RxWord[ConvWordIndex]);
    END_IF;
END_FOR;

ConvUnitOK := (RCON2_SpeedUnit_mm_s = LREAL#1.0) OR
              (RCON2_SpeedUnit_mm_s = LREAL#0.1);

// 【①-2 共通状態】IN00はユニット全体、IN01は各軸のリンク情報です。
// TestABit(ワード, bit番号)は、そのスイッチがONかをBOOLで取り出す命令です。
// 例：IN01のb0は軸No.0→配列[1]、b1は軸No.1→配列[2]。配列番号と実機軸番号は1違います。
// 共通固定領域。ここで使うbit番号は取説の論理bitです（MJ0384 6-24～6-25）。
RCON2_GwRun := TestABit(RCON2_RxWord[0], USINT#15);
RCON2_GwControllerCommLatch := TestABit(RCON2_RxWord[0], USINT#14);
RCON2_GwAxisCommError := TestABit(RCON2_RxWord[0], USINT#13);
RCON2_GwManual := TestABit(RCON2_RxWord[0], USINT#12);
RCON2_GwHeavyAlarm := TestABit(RCON2_RxWord[0], USINT#11);
RCON2_GwLightAlarm := TestABit(RCON2_RxWord[0], USINT#10);
RCON2_GwSystemStop := TestABit(RCON2_RxWord[0], USINT#8);
RCON2_GwAlarmCode := WORD_TO_UINT(RCON2_RxWord[0] AND WORD#16#00FF);
FOR ConvWordIndex := INT#0 TO INT#4 DO
    RCON2_PowerStateRaw[ConvWordIndex] := RCON2_RxWord[ConvWordIndex + INT#2];
END_FOR;

// 【①-3 軸ごとに同じ読取りを繰り返す】
// FORは1～5軸を順番に処理します。ConvBaseはその軸の先頭番号です。
// 計算：8+(軸番号-1)×8。1軸目=8、2軸目=16、3軸目=24。先頭8ワードは共通領域です。
FOR ConvAxisIndex := INT#1 TO INT#5 DO
    ConvBase := INT#8 + (ConvAxisIndex - INT#1) * INT#8;
    RCON2_AxisLinked[ConvAxisIndex] :=
        TestABit(RCON2_RxWord[1], INT_TO_USINT(ConvAxisIndex - INT#1));

// 例：下位2540／上位0なら32bit値2540→25.40mm。
// 上位を16bit左に動かして下位とORで重ねます。SHLが左シフト、ORがビットの合成です。
// 負位置はDWORD_TO_DINTで符号を復元。下位62996／上位65535なら-2540→-25.40mm。
    // 現在位置：下位・上位を結合、符号付き32bitとして解釈、0.01mmをmmへ。
    ConvDWord := SHL(WORD_TO_DWORD(RCON2_RxWord[ConvBase + INT#1]), ULINT#16)
                 OR WORD_TO_DWORD(RCON2_RxWord[ConvBase]);
    RCON2_IN[ConvAxisIndex].ActualPos_mm :=
        DINT_TO_LREAL(DWORD_TO_DINT(ConvDWord)) * LREAL#0.01;

    // 電流：32bitのmA。RCON-PCでは指令電流であり、実測トルクではありません。
    ConvDWord := SHL(WORD_TO_DWORD(RCON2_RxWord[ConvBase + INT#3]), ULINT#16)
                 OR WORD_TO_DWORD(RCON2_RxWord[ConvBase + INT#2]);
    RCON2_IN[ConvAxisIndex].Current_mA := DWORD_TO_DINT(ConvDWord);

    // 現在速度：16bitの負数をINTとして読む。UINTのまま速度にしません。
    IF ConvUnitOK THEN
        RCON2_IN[ConvAxisIndex].ActualSpeed_mm_s :=
            INT_TO_LREAL(WORD_TO_INT(RCON2_RxWord[ConvBase + INT#4])) * RCON2_SpeedUnit_mm_s;
    END_IF;
    // 単位不明のとき速度は前値を保持し、DataValidはFALSEにします。
    // 軸内の+5ワードは予約のため値を使用しません。
    RCON2_IN[ConvAxisIndex].AlarmCode := WORD_TO_UINT(RCON2_RxWord[ConvBase + INT#6]);

// 例：Status.ServoReady=TRUEは「サーボON状態を受信した」という意味。
// OUT側Control.ServoOn=TRUEは「サーボONを要求する」という意味で、指令と結果を区別します。
    // 状態ワード：12個のBOOLへ分解。予約b6,b9～11は使いません。
    RCON2_IN[ConvAxisIndex].Status.PositionDone := TestABit(RCON2_RxWord[ConvBase + INT#7], USINT#0);
    RCON2_IN[ConvAxisIndex].Status.HomeDone := TestABit(RCON2_RxWord[ConvBase + INT#7], USINT#1);
    RCON2_IN[ConvAxisIndex].Status.Moving := TestABit(RCON2_RxWord[ConvBase + INT#7], USINT#2);
    RCON2_IN[ConvAxisIndex].Status.Alarm := TestABit(RCON2_RxWord[ConvBase + INT#7], USINT#3);
    RCON2_IN[ConvAxisIndex].Status.ServoReady := TestABit(RCON2_RxWord[ConvBase + INT#7], USINT#4);
    RCON2_IN[ConvAxisIndex].Status.PushMiss := TestABit(RCON2_RxWord[ConvBase + INT#7], USINT#5);
    RCON2_IN[ConvAxisIndex].Status.OverloadWarning := TestABit(RCON2_RxWord[ConvBase + INT#7], USINT#7);
    RCON2_IN[ConvAxisIndex].Status.CommandDone := TestABit(RCON2_RxWord[ConvBase + INT#7], USINT#8);
    RCON2_IN[ConvAxisIndex].Status.Zone1 := TestABit(RCON2_RxWord[ConvBase + INT#7], USINT#12);
    RCON2_IN[ConvAxisIndex].Status.Zone2 := TestABit(RCON2_RxWord[ConvBase + INT#7], USINT#13);
    RCON2_IN[ConvAxisIndex].Status.ControllerReady := TestABit(RCON2_RxWord[ConvBase + INT#7], USINT#14);
    RCON2_IN[ConvAxisIndex].Status.EmergencyStop := TestABit(RCON2_RxWord[ConvBase + INT#7], USINT#15);

    // DataValidは直接受信bitではなく、今回の内部設計で決めた内部判定です。
    // CommOKはCPUの実通信状態から別途作成。単にTRUE固定にしないでください。
    // DataValidは運転許可や安全保証ではありません。各異常・原点等は別途確認。
    RCON2_IN[ConvAxisIndex].DataValid := RCON2_CommOK AND RCON2_LayoutConfirmed
        AND RCON2_ByteOrderConfirmed AND ConvUnitOK AND RCON2_GwRun
        AND RCON2_AxisLinked[ConvAxisIndex] AND NOT RCON2_GwAxisCommError;
END_FOR;

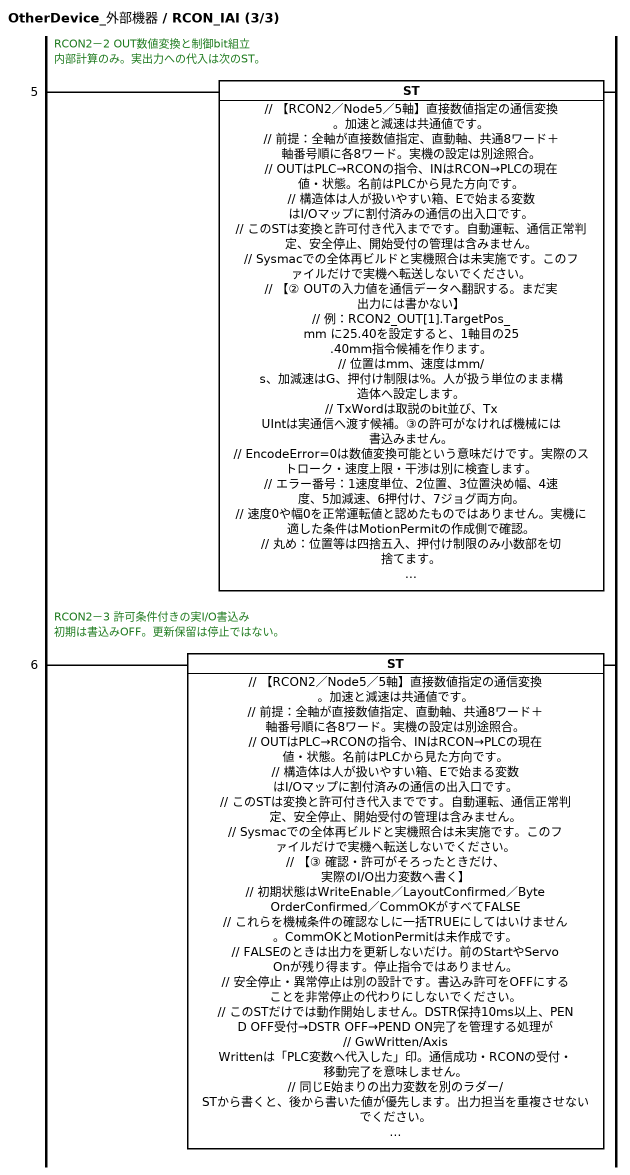
(* Rung 5: RCON2－2 OUT数値変換と制御bit組立 / 内部計算のみ。実出力への代入は次のST。 *)
// 【RCON2／Node5／5軸】直接数値指定の通信変換。加速と減速は共通値です。
// 前提：全軸が直接数値指定、直動軸、共通8ワード＋軸番号順に各8ワード。実機の設定は別途照合。
// OUTはPLC→RCONの指令、INはRCON→PLCの現在値・状態。名前はPLCから見た方向です。
// 構造体は人が扱いやすい箱、Eで始まる変数はI/Oマップに割付済みの通信の出入口です。
// このSTは変換と許可付き代入までです。自動運転、通信正常判定、安全停止、開始受付の管理は含みません。
// Sysmacでの全体再ビルドと実機照合は未実施です。このファイルだけで実機へ転送しないでください。
// 【② OUTの入力値を通信データへ翻訳する。まだ実出力には書かない】
// 例：RCON2_OUT[1].TargetPos_mm に25.40を設定すると、1軸目の25.40mm指令候補を作ります。
// 位置はmm、速度はmm/s、加減速はG、押付け制限は%。人が扱う単位のまま構造体へ設定します。
// TxWordは取説のbit並び、TxUIntは実通信へ渡す候補。③の許可がなければ機械には書込みません。
// EncodeError=0は数値変換可能という意味だけです。実際のストローク・速度上限・干渉は別に検査します。
// エラー番号：1速度単位、2位置、3位置決め幅、4速度、5加減速、6押付け、7ジョグ両方向。
// 速度0や幅0を正常運転値と認めたものではありません。実機に適した条件はMotionPermitの作成側で確認。
// 丸め：位置等は四捨五入、押付け制限のみ小数部を切捨てます。

ConvUnitOK := (RCON2_SpeedUnit_mm_s = LREAL#1.0) OR
              (RCON2_SpeedUnit_mm_s = LREAL#0.1);

// 共通制御：MONは論理b15、RTEは論理b13。他のbitは0。
// MONを落とす処理を安全停止として扱わないでください。
RCON2_TxWord[0] := WORD#16#0000;
IF RCON2_GwMON_Request THEN
    RCON2_TxWord[0] := RCON2_TxWord[0] OR WORD#16#8000;
END_IF;
IF RCON2_GwRTE_Request THEN
    RCON2_TxWord[0] := RCON2_TxWord[0] OR WORD#16#2000;
END_IF;

FOR ConvAxisIndex := INT#1 TO INT#5 DO
    ConvBase := INT#8 + (ConvAxisIndex - INT#1) * INT#8;
    RCON2_EncodeError[ConvAxisIndex] := UINT#0;

    // 比較で範囲を確認してから型変換するため、NaN・無限大も変換対象から外れます。
    // 位置・幅9999.99mmはこの案で採用する通信範囲の上限で、実機ストロークではありません。
    IF NOT ConvUnitOK THEN
        RCON2_EncodeError[ConvAxisIndex] := UINT#1;
    ELSIF NOT ((RCON2_OUT[ConvAxisIndex].TargetPos_mm >= LREAL#-9999.99) AND
               (RCON2_OUT[ConvAxisIndex].TargetPos_mm <= LREAL#9999.99)) THEN
        RCON2_EncodeError[ConvAxisIndex] := UINT#2;
    ELSIF NOT ((RCON2_OUT[ConvAxisIndex].PositionBand_mm >= LREAL#0.0) AND
               (RCON2_OUT[ConvAxisIndex].PositionBand_mm <= LREAL#9999.99)) THEN
        RCON2_EncodeError[ConvAxisIndex] := UINT#3;
    ELSIF NOT ((RCON2_OUT[ConvAxisIndex].Speed_mm_s >= LREAL#0.0) AND
               (RCON2_OUT[ConvAxisIndex].Speed_mm_s <= LREAL#65535.0 * RCON2_SpeedUnit_mm_s)) THEN
        RCON2_EncodeError[ConvAxisIndex] := UINT#4;
    ELSIF NOT ((RCON2_OUT[ConvAxisIndex].AccDec_G >= LREAL#0.0) AND
               (RCON2_OUT[ConvAxisIndex].AccDec_G <= LREAL#655.35)) THEN
        RCON2_EncodeError[ConvAxisIndex] := UINT#5;
    ELSIF NOT ((RCON2_OUT[ConvAxisIndex].PushLimit_pct >= LREAL#0.0) AND
               (RCON2_OUT[ConvAxisIndex].PushLimit_pct <= LREAL#200.0)) THEN
        RCON2_EncodeError[ConvAxisIndex] := UINT#6;
    ELSIF RCON2_OUT[ConvAxisIndex].Control.JogMinus AND RCON2_OUT[ConvAxisIndex].Control.JogPlus THEN
        RCON2_EncodeError[ConvAxisIndex] := UINT#7;
    END_IF;

    RCON2_EncodeOK[ConvAxisIndex] := RCON2_EncodeError[ConvAxisIndex] = UINT#0;
    IF RCON2_EncodeOK[ConvAxisIndex] THEN
    // 【数値例】TargetPos_mm=25.40→×100で2540。下位ワード2540、上位ワード0。
// 700.25mm→70025なので下位4489、上位1。65536を超えた分が上位に入ります。
// DINTは符号付きの数、DWORDは同じ32bitの模様。負数の符号を壊さず分割するために使い分けます。
// TRUNCは小数部を捨てます。正数+0.5／負数-0.5を先に行い、四捨五入を明示しています。
    // 目標位置：mmから0.01mmの符号付き整数へ。
        ConvScaled := RCON2_OUT[ConvAxisIndex].TargetPos_mm * LREAL#100.0;
        IF ConvScaled >= LREAL#0.0 THEN
            ConvPos := LINT_TO_DINT(TRUNC(ConvScaled + LREAL#0.5));
        ELSE
            ConvPos := LINT_TO_DINT(TRUNC(ConvScaled - LREAL#0.5));
        END_IF;
        // 負数を含む32bitパターンを保ち、下位・上位の16bitへ分割。
        ConvDWord := DINT_TO_DWORD(ConvPos);
        RCON2_TxWord[ConvBase] := DWORD_TO_WORD(ConvDWord AND DWORD#16#0000FFFF);
        RCON2_TxWord[ConvBase + INT#1] := DWORD_TO_WORD(SHR(ConvDWord, ULINT#16));

        // 位置決め幅：非負の内部整数としてUDINTを選定（メーカーの符号なし保証ではありません）。
        ConvBand := LINT_TO_UDINT(TRUNC(RCON2_OUT[ConvAxisIndex].PositionBand_mm * LREAL#100.0 + LREAL#0.5));
        ConvDWord := UDINT_TO_DWORD(ConvBand);
        RCON2_TxWord[ConvBase + INT#2] := DWORD_TO_WORD(ConvDWord AND DWORD#16#0000FFFF);
        RCON2_TxWord[ConvBase + INT#3] := DWORD_TO_WORD(SHR(ConvDWord, ULINT#16));

// 速度20mm/s：速度単位1.0なら20、0.1なら200を送信します。
// 加減速0.20G：×100して20。加速と減速の両方に同じ値を使います。
// 押付け50%：×255÷100=127.5を切捨てて127。押付けの使用可否・上限は実機仕様で別確認。
        // 速度は1カウント量が1.0か0.1かで値が10倍変わります。
        ConvSpeed := LINT_TO_UINT(TRUNC(RCON2_OUT[ConvAxisIndex].Speed_mm_s / RCON2_SpeedUnit_mm_s + LREAL#0.5));
        ConvAccDec := LINT_TO_UINT(TRUNC(RCON2_OUT[ConvAxisIndex].AccDec_G * LREAL#100.0 + LREAL#0.5));
        ConvPush := LINT_TO_UINT(TRUNC(RCON2_OUT[ConvAxisIndex].PushLimit_pct * LREAL#255.0 / LREAL#100.0));
        RCON2_TxWord[ConvBase + INT#4] := UINT_TO_WORD(ConvSpeed);
        RCON2_TxWord[ConvBase + INT#5] := UINT_TO_WORD(ConvAccDec);
        RCON2_TxWord[ConvBase + INT#6] := UINT_TO_WORD(ConvPush);
    END_IF;
    // 不正値の場合、数値ワードは前値保持。EncodeOK=FALSEで03の書込みを抑止。
    // 前値保持は停止指令ではありません。停止・異常処理は別途設計してください。

    // Controlを論理bitへ詰める。予約b9は必ず0。
    RCON2_TxWord[ConvBase + INT#7] := WORD#16#0000;
// b0 DSTR／Control.Start：TRUEで開始要求。受付応答と10ms以上の保持を確認してOFF。常時ONにしない。
    IF RCON2_OUT[ConvAxisIndex].Control.Start THEN
        RCON2_TxWord[ConvBase + INT#7] := RCON2_TxWord[ConvBase + INT#7] OR WORD#16#0001;
    END_IF;
// b1 HOME／Control.Home：TRUEで原点復帰を指令。原点復帰完了はIN側HomeDoneで確認。
    IF RCON2_OUT[ConvAxisIndex].Control.Home THEN
        RCON2_TxWord[ConvBase + INT#7] := RCON2_TxWord[ConvBase + INT#7] OR WORD#16#0002;
    END_IF;
// b2 STP／Control.Pause：TRUEで一時停止、FALSEで解除。非常停止・安全停止の代用ではない。
    IF RCON2_OUT[ConvAxisIndex].Control.Pause THEN
        RCON2_TxWord[ConvBase + INT#7] := RCON2_TxWord[ConvBase + INT#7] OR WORD#16#0004;
    END_IF;
// b3 RES／Control.Reset：TRUEでアラームリセット要求。コールドスタート級の異常には使用できない。
    IF RCON2_OUT[ConvAxisIndex].Control.Reset THEN
        RCON2_TxWord[ConvBase + INT#7] := RCON2_TxWord[ConvBase + INT#7] OR WORD#16#0008;
    END_IF;
// b4 SON／Control.ServoOn：TRUEでサーボON要求。ON状態はIN側ServoReadyで確認。
    IF RCON2_OUT[ConvAxisIndex].Control.ServoOn THEN
        RCON2_TxWord[ConvBase + INT#7] := RCON2_TxWord[ConvBase + INT#7] OR WORD#16#0010;
    END_IF;
// b5 JISL／Control.InchingSelect：TRUEは一定距離のインチング、FALSEは押している間のジョグ。
    IF RCON2_OUT[ConvAxisIndex].Control.InchingSelect THEN
        RCON2_TxWord[ConvBase + INT#7] := RCON2_TxWord[ConvBase + INT#7] OR WORD#16#0020;
    END_IF;
// b6 JVEL／Control.JogSpeedSelect：FALSEは速度No.26・距離No.48、TRUEは速度No.47または指令速度・距離No.49。
    IF RCON2_OUT[ConvAxisIndex].Control.JogSpeedSelect THEN
        RCON2_TxWord[ConvBase + INT#7] := RCON2_TxWord[ConvBase + INT#7] OR WORD#16#0040;
    END_IF;
// b7 JOG-／Control.JogMinus：TRUEで原点方向へジョグ。反対方向指令との同時ONを防ぐ。
    IF RCON2_OUT[ConvAxisIndex].Control.JogMinus THEN
        RCON2_TxWord[ConvBase + INT#7] := RCON2_TxWord[ConvBase + INT#7] OR WORD#16#0080;
    END_IF;
// b8 JOG+／Control.JogPlus：TRUEで反原点方向へジョグ。反対方向指令との同時ONを防ぐ。
    IF RCON2_OUT[ConvAxisIndex].Control.JogPlus THEN
        RCON2_TxWord[ConvBase + INT#7] := RCON2_TxWord[ConvBase + INT#7] OR WORD#16#0100;
    END_IF;
// b10 GSL0／Control.GainSelect0：GainSelect1と組合せてサーボゲインセット0～3を選ぶ。機械調整用。
    IF RCON2_OUT[ConvAxisIndex].Control.GainSelect0 THEN
        RCON2_TxWord[ConvBase + INT#7] := RCON2_TxWord[ConvBase + INT#7] OR WORD#16#0400;
    END_IF;
// b11 GSL1／Control.GainSelect1：GainSelect0との2bitで選択。速度指令とは別の機能。
    IF RCON2_OUT[ConvAxisIndex].Control.GainSelect1 THEN
        RCON2_TxWord[ConvBase + INT#7] := RCON2_TxWord[ConvBase + INT#7] OR WORD#16#0800;
    END_IF;
// b12 PUSH／Control.PushEnable：TRUEは押付け、FALSEは通常位置決め。押付け条件は別途確認。
    IF RCON2_OUT[ConvAxisIndex].Control.PushEnable THEN
        RCON2_TxWord[ConvBase + INT#7] := RCON2_TxWord[ConvBase + INT#7] OR WORD#16#1000;
    END_IF;
// b13 DIR／Control.PushDirection：CON方式押付け時、TRUEは反原点方向、FALSEは原点方向。
    IF RCON2_OUT[ConvAxisIndex].Control.PushDirection THEN
        RCON2_TxWord[ConvBase + INT#7] := RCON2_TxWord[ConvBase + INT#7] OR WORD#16#2000;
    END_IF;
// b14 INC／Control.RelativeMove：FALSEは絶対座標、TRUEは現在位置からの相対移動量。
    IF RCON2_OUT[ConvAxisIndex].Control.RelativeMove THEN
        RCON2_TxWord[ConvBase + INT#7] := RCON2_TxWord[ConvBase + INT#7] OR WORD#16#4000;
    END_IF;
// b15 BKRL／Control.BrakeRelease：TRUEはブレーキ強制解除。通常FALSE。縦軸では落下等の危険がある。
    IF RCON2_OUT[ConvAxisIndex].Control.BrakeRelease THEN
        RCON2_TxWord[ConvBase + INT#7] := RCON2_TxWord[ConvBase + INT#7] OR WORD#16#8000;
    END_IF;
END_FOR;

// 論理ワードから実際に送るUINTへ。INと同じ1ワード内のバイト交換を適用します。
FOR ConvWordIndex := INT#0 TO INT#47 DO
    ConvWord := RCON2_TxWord[ConvWordIndex];
    IF RCON2_SwapBytes THEN
        ConvWord := Swap(ConvWord);
    END_IF;
    RCON2_TxUInt[ConvWordIndex] := WORD_TO_UINT(ConvWord);
END_FOR;
(* Rung 6: RCON2－3 許可条件付きの実I/O書込み / 初期は書込みOFF。更新保留は停止ではない。 *)
// 【RCON2／Node5／5軸】直接数値指定の通信変換。加速と減速は共通値です。
// 前提：全軸が直接数値指定、直動軸、共通8ワード＋軸番号順に各8ワード。実機の設定は別途照合。
// OUTはPLC→RCONの指令、INはRCON→PLCの現在値・状態。名前はPLCから見た方向です。
// 構造体は人が扱いやすい箱、Eで始まる変数はI/Oマップに割付済みの通信の出入口です。
// このSTは変換と許可付き代入までです。自動運転、通信正常判定、安全停止、開始受付の管理は含みません。
// Sysmacでの全体再ビルドと実機照合は未実施です。このファイルだけで実機へ転送しないでください。
// 【③ 確認・許可がそろったときだけ、実際のI/O出力変数へ書く】
// 初期状態はWriteEnable／LayoutConfirmed／ByteOrderConfirmed／CommOKがすべてFALSEです。
// これらを機械条件の確認なしに一括TRUEにしてはいけません。CommOKとMotionPermitは未作成です。
// FALSEのときは出力を更新しないだけ。前のStartやServoOnが残り得ます。停止指令ではありません。
// 安全停止・異常停止は別の設計です。書込み許可をOFFにすることを非常停止の代わりにしないでください。
// このSTだけでは動作開始しません。DSTR保持10ms以上、PEND OFF受付→DSTR OFF→PEND ON完了を管理する処理が必要です。
// GwWritten/AxisWrittenは「PLC変数へ代入した」印。通信成功・RCONの受付・移動完了を意味しません。
// 同じE始まりの出力変数を別のラダー/STから書くと、後から書いた値が優先します。出力担当を重複させないでください。

RCON2_GwWritten := FALSE;
FOR ConvAxisIndex := INT#1 TO INT#5 DO
    RCON2_AxisWritten[ConvAxisIndex] := FALSE;
END_FOR;

IF RCON2_WriteEnable AND RCON2_LayoutConfirmed AND RCON2_ByteOrderConfirmed AND RCON2_CommOK THEN
// 共通指令はMON/RTEのみ。最初のRUN応答に必要なため、軸DataValidとは別にGwApplyで許可します。
    IF RCON2_GwApply THEN
        E005_Out_OUT00_2003_01_1 := RCON2_TxUInt[0];
        RCON2_GwWritten := TRUE;
    END_IF;

// 1軸目＝実機軸No.0。OUT08～OUT15の8ワードをまとめて代入。
// AxisApply=この軸の更新許可、EncodeOK=変換OK、DataValid=入力情報の条件確認、MotionPermit=機械側の運転許可。
// 途中1ワードだけではなく、位置・幅・速度・加減速・押付け・制御を一組として渡します。
    IF RCON2_AxisApply[1] AND RCON2_EncodeOK[1] AND RCON2_IN[1].DataValid
       AND RCON2_MotionPermit[1] THEN
        E005_Out_OUT08_2003_09_1 := RCON2_TxUInt[8];
        E005_Out_OUT09_2003_0A_1 := RCON2_TxUInt[9];
        E005_Out_OUT10_2003_0B_1 := RCON2_TxUInt[10];
        E005_Out_OUT11_2003_0C_1 := RCON2_TxUInt[11];
        E005_Out_OUT12_2003_0D_1 := RCON2_TxUInt[12];
        E005_Out_OUT13_2003_0E_1 := RCON2_TxUInt[13];
        E005_Out_OUT14_2003_0F_1 := RCON2_TxUInt[14];
        E005_Out_OUT15_2003_10_1 := RCON2_TxUInt[15];
        RCON2_AxisWritten[1] := TRUE;
    END_IF;

// 2軸目＝実機軸No.1。OUT16～OUT23の8ワードをまとめて代入。
// AxisApply=この軸の更新許可、EncodeOK=変換OK、DataValid=入力情報の条件確認、MotionPermit=機械側の運転許可。
// 途中1ワードだけではなく、位置・幅・速度・加減速・押付け・制御を一組として渡します。
    IF RCON2_AxisApply[2] AND RCON2_EncodeOK[2] AND RCON2_IN[2].DataValid
       AND RCON2_MotionPermit[2] THEN
        E005_Out_OUT16_2003_11_1 := RCON2_TxUInt[16];
        E005_Out_OUT17_2003_12_1 := RCON2_TxUInt[17];
        E005_Out_OUT18_2003_13_1 := RCON2_TxUInt[18];
        E005_Out_OUT19_2003_14_1 := RCON2_TxUInt[19];
        E005_Out_OUT20_2003_15_1 := RCON2_TxUInt[20];
        E005_Out_OUT21_2003_16_1 := RCON2_TxUInt[21];
        E005_Out_OUT22_2003_17_1 := RCON2_TxUInt[22];
        E005_Out_OUT23_2003_18_1 := RCON2_TxUInt[23];
        RCON2_AxisWritten[2] := TRUE;
    END_IF;

// 3軸目＝実機軸No.2。OUT24～OUT31の8ワードをまとめて代入。
// AxisApply=この軸の更新許可、EncodeOK=変換OK、DataValid=入力情報の条件確認、MotionPermit=機械側の運転許可。
// 途中1ワードだけではなく、位置・幅・速度・加減速・押付け・制御を一組として渡します。
    IF RCON2_AxisApply[3] AND RCON2_EncodeOK[3] AND RCON2_IN[3].DataValid
       AND RCON2_MotionPermit[3] THEN
        E005_Out_OUT24_2003_19_1 := RCON2_TxUInt[24];
        E005_Out_OUT25_2003_1A_1 := RCON2_TxUInt[25];
        E005_Out_OUT26_2003_1B_1 := RCON2_TxUInt[26];
        E005_Out_OUT27_2003_1C_1 := RCON2_TxUInt[27];
        E005_Out_OUT28_2003_1D_1 := RCON2_TxUInt[28];
        E005_Out_OUT29_2003_1E_1 := RCON2_TxUInt[29];
        E005_Out_OUT30_2003_1F_1 := RCON2_TxUInt[30];
        E005_Out_OUT31_2003_20_1 := RCON2_TxUInt[31];
        RCON2_AxisWritten[3] := TRUE;
    END_IF;

// 4軸目＝実機軸No.3。OUT32～OUT39の8ワードをまとめて代入。
// AxisApply=この軸の更新許可、EncodeOK=変換OK、DataValid=入力情報の条件確認、MotionPermit=機械側の運転許可。
// 途中1ワードだけではなく、位置・幅・速度・加減速・押付け・制御を一組として渡します。
    IF RCON2_AxisApply[4] AND RCON2_EncodeOK[4] AND RCON2_IN[4].DataValid
       AND RCON2_MotionPermit[4] THEN
        E005_Out_OUT32_2003_21_1 := RCON2_TxUInt[32];
        E005_Out_OUT33_2003_22_1 := RCON2_TxUInt[33];
        E005_Out_OUT34_2003_23_1 := RCON2_TxUInt[34];
        E005_Out_OUT35_2003_24_1 := RCON2_TxUInt[35];
        E005_Out_OUT36_2003_25_1 := RCON2_TxUInt[36];
        E005_Out_OUT37_2003_26_1 := RCON2_TxUInt[37];
        E005_Out_OUT38_2003_27_1 := RCON2_TxUInt[38];
        E005_Out_OUT39_2003_28_1 := RCON2_TxUInt[39];
        RCON2_AxisWritten[4] := TRUE;
    END_IF;

// 5軸目＝実機軸No.4。OUT40～OUT47の8ワードをまとめて代入。
// AxisApply=この軸の更新許可、EncodeOK=変換OK、DataValid=入力情報の条件確認、MotionPermit=機械側の運転許可。
// 途中1ワードだけではなく、位置・幅・速度・加減速・押付け・制御を一組として渡します。
    IF RCON2_AxisApply[5] AND RCON2_EncodeOK[5] AND RCON2_IN[5].DataValid
       AND RCON2_MotionPermit[5] THEN
        E005_Out_OUT40_2003_29_1 := RCON2_TxUInt[40];
        E005_Out_OUT41_2003_2A_1 := RCON2_TxUInt[41];
        E005_Out_OUT42_2003_2B_1 := RCON2_TxUInt[42];
        E005_Out_OUT43_2003_2C_1 := RCON2_TxUInt[43];
        E005_Out_OUT44_2003_2D_1 := RCON2_TxUInt[44];
        E005_Out_OUT45_2003_2E_1 := RCON2_TxUInt[45];
        E005_Out_OUT46_2003_2F_1 := RCON2_TxUInt[46];
        E005_Out_OUT47_2003_30_1 := RCON2_TxUInt[47];
        RCON2_AxisWritten[5] := TRUE;
    END_IF;
END_IF;
// OUT01～07、OUT48～55は、このSTからは一切書き換えません。
// 現在の実機設定・別処理の用途が未確認なので、余剰領域を勝手にゼロクリアしません。

(* Section DLEP1_GT2: ladder, written here as Structured Text *)

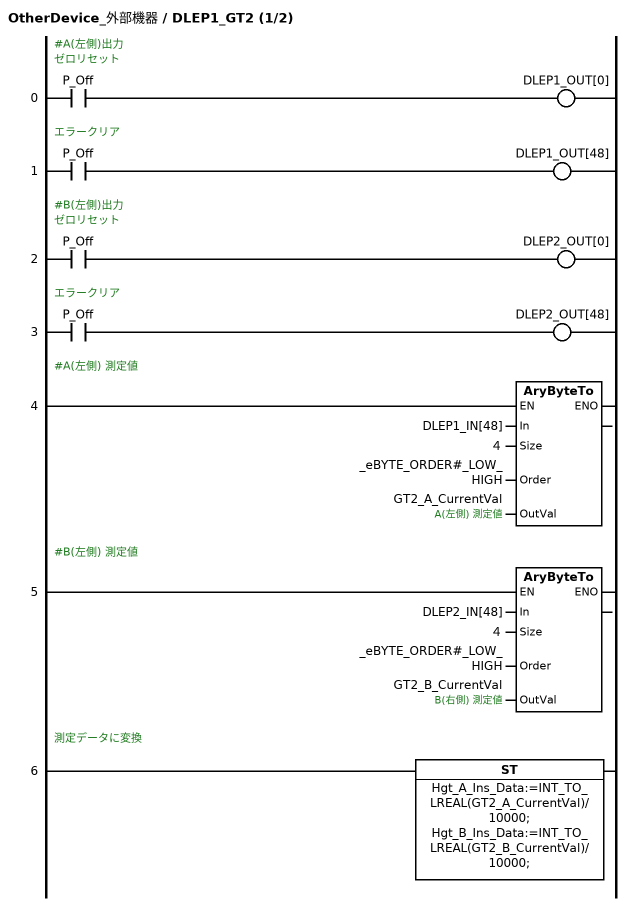
(* Rung 0: #A(左側)出力 / ゼロリセット *)
DLEP1_OUT[0] := P_Off;
(* Rung 1: エラークリア *)
DLEP1_OUT[48] := P_Off;
(* Rung 2: #B(左側)出力 / ゼロリセット *)
DLEP2_OUT[0] := P_Off;
(* Rung 3: エラークリア *)
DLEP2_OUT[48] := P_Off;
(* Rung 4: #A(左側) 測定値 *)
AryByteTo(In := DLEP1_IN[48], Size := ４, Order := _eBYTE_ORDER#_LOW_HIGH, OutVal := GT2_A_CurrentVal);
(* Rung 5: #B(左側) 測定値 *)
AryByteTo(In := DLEP2_IN[48], Size := ４, Order := _eBYTE_ORDER#_LOW_HIGH, OutVal := GT2_B_CurrentVal);
(* Rung 6: 測定データに変換 *)
Hgt_A_Ins_Data:=INT_TO_LREAL(GT2_A_CurrentVal)/10000;
Hgt_B_Ins_Data:=INT_TO_LREAL(GT2_B_CurrentVal)/10000;

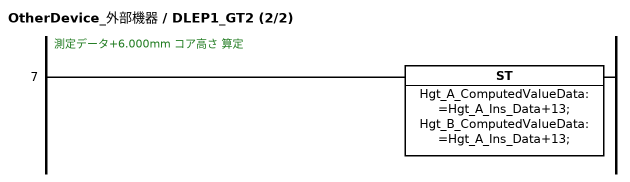
(* Rung 7: 測定データ+6.000mm コア高さ 算定 *)
Hgt_A_ComputedValueData:=Hgt_A_Ins_Data+13;
Hgt_B_ComputedValueData:=Hgt_A_Ins_Data+13;

(* Section FH_5552_10: ladder, written here as Structured Text *)

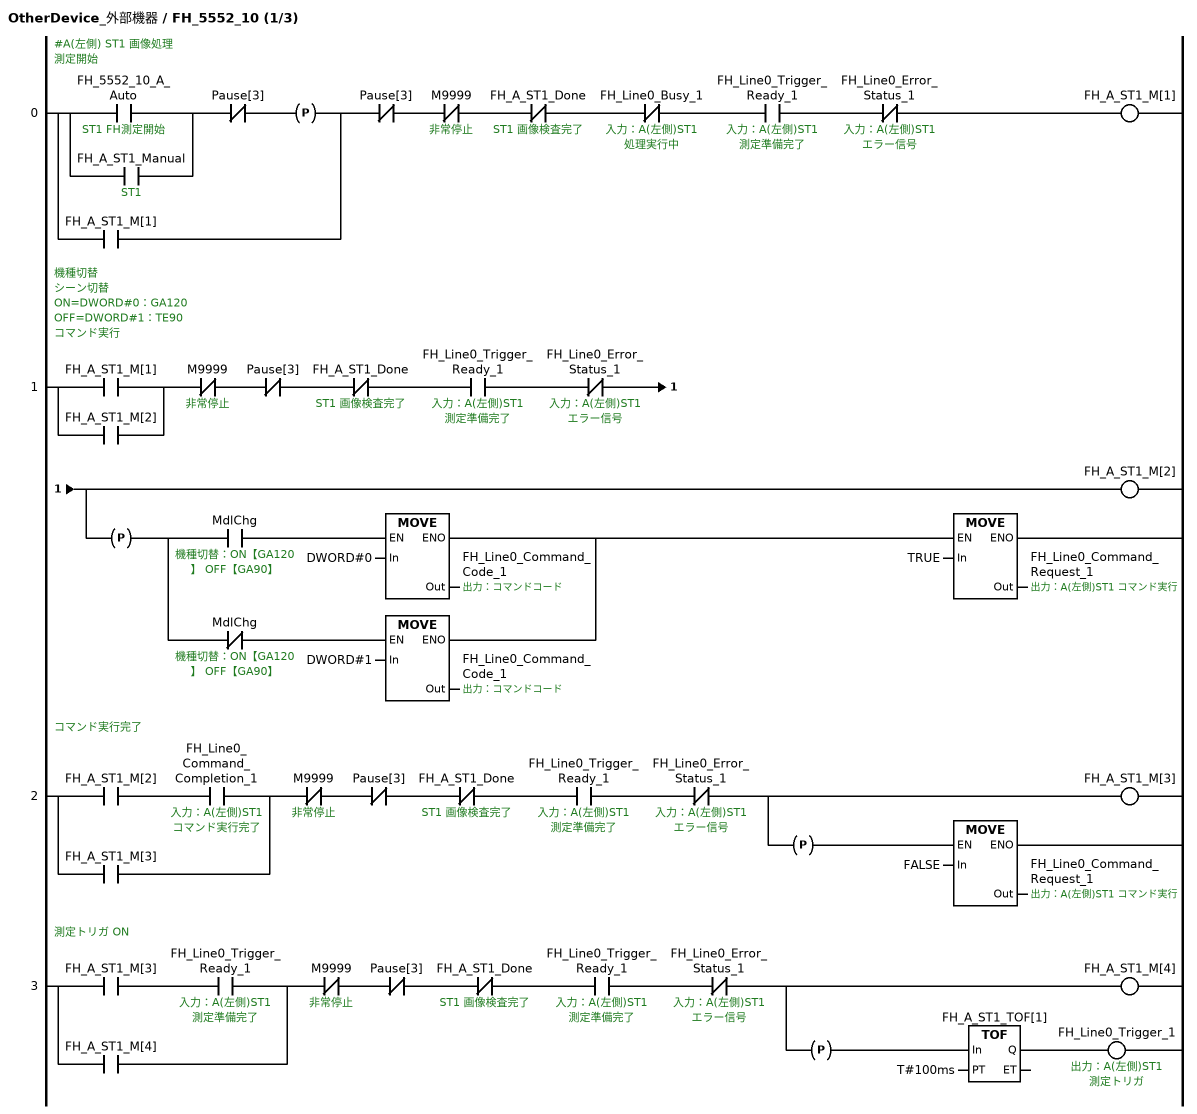
(* Rung 0: #A(左側) ST1 画像処理 / 測定開始 *)
_e1(CLK := (FH_5552_10_A_Auto OR FH_A_ST1_Manual) AND NOT Pause[3]);
FH_A_ST1_M[1] := (_e1.Q OR FH_A_ST1_M[1]) AND NOT Pause[3] AND NOT M9999 AND NOT FH_A_ST1_Done AND NOT FH_Line0_Busy_1 AND FH_Line0_Trigger_Ready_1 AND NOT FH_Line0_Error_Status_1;
(* Rung 1: 機種切替 / シーン切替 / ON=DWORD#0：GA120 / OFF=DWORD#1：TE90 / コマンド実行 *)
_p2 := (FH_A_ST1_M[1] OR FH_A_ST1_M[2]) AND NOT M9999 AND NOT Pause[3] AND NOT FH_A_ST1_Done AND FH_Line0_Trigger_Ready_1 AND NOT FH_Line0_Error_Status_1;
FH_A_ST1_M[2] := _p2;
_e3(CLK := _p2);
IF _e3.Q AND MdlChg THEN FH_Line0_Command_Code_1 := DWORD#0; END_IF;
IF _e3.Q AND NOT MdlChg THEN FH_Line0_Command_Code_1 := DWORD#1; END_IF;
IF _e3.Q AND (MdlChg OR NOT MdlChg) THEN FH_Line0_Command_Request_1 := TRUE; END_IF;
(* Rung 2: コマンド実行完了 *)
_p4 := ((FH_A_ST1_M[2] AND FH_Line0_Command_Completion_1) OR FH_A_ST1_M[3]) AND NOT M9999 AND NOT Pause[3] AND NOT FH_A_ST1_Done AND FH_Line0_Trigger_Ready_1 AND NOT FH_Line0_Error_Status_1;
FH_A_ST1_M[3] := _p4;
_e5(CLK := _p4);
IF _e5.Q THEN FH_Line0_Command_Request_1 := FALSE; END_IF;
(* Rung 3: 測定トリガ ON *)
_p6 := ((FH_A_ST1_M[3] AND FH_Line0_Trigger_Ready_1) OR FH_A_ST1_M[4]) AND NOT M9999 AND NOT Pause[3] AND NOT FH_A_ST1_Done AND FH_Line0_Trigger_Ready_1 AND NOT FH_Line0_Error_Status_1;
FH_A_ST1_M[4] := _p6;
_e7(CLK := _p6);
FH_A_ST1_TOF[1](In := _e7.Q, PT := T#100ms);
FH_Line0_Trigger_1 := FH_A_ST1_TOF[1].Q;

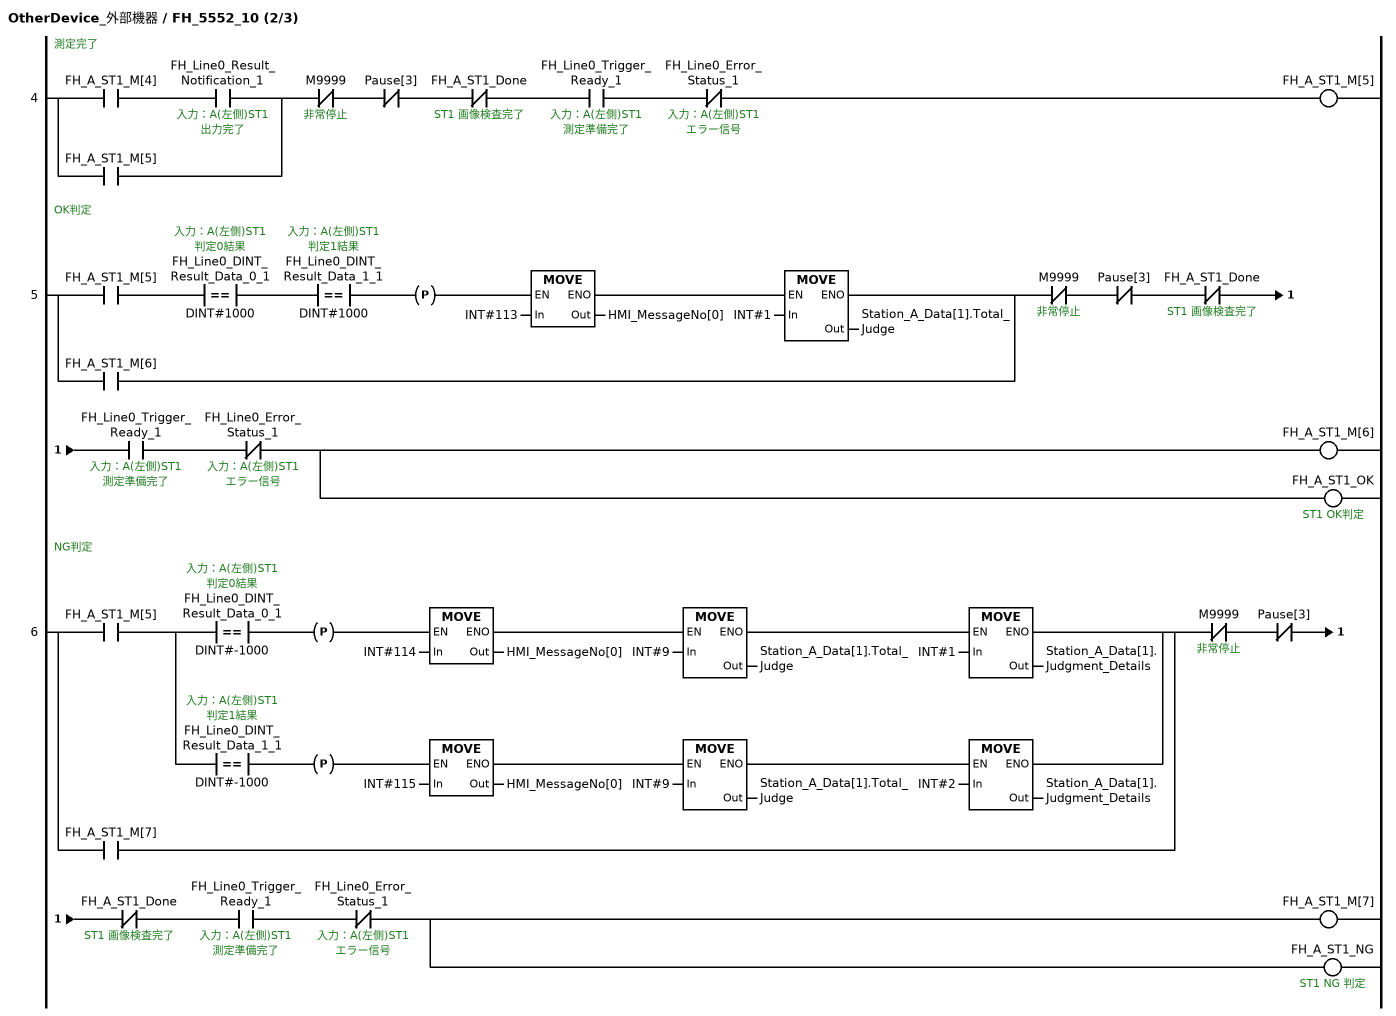
(* Rung 4: 測定完了 *)
FH_A_ST1_M[5] := ((FH_A_ST1_M[4] AND FH_Line0_Result_Notification_1) OR FH_A_ST1_M[5]) AND NOT M9999 AND NOT Pause[3] AND NOT FH_A_ST1_Done AND FH_Line0_Trigger_Ready_1 AND NOT FH_Line0_Error_Status_1;
(* Rung 5: OK判定 *)
_e8(CLK := FH_A_ST1_M[5] AND (FH_Line0_DINT_Result_Data_0_1 = DINT#1000) AND (FH_Line0_DINT_Result_Data_1_1 = DINT#1000));
IF _e8.Q THEN
    HMI_MessageNo[0] := INT#113;
    Station_A_Data[1].Total_Judge := INT#1;
END_IF;
_p9 := (_e8.Q OR FH_A_ST1_M[6]) AND NOT M9999 AND NOT Pause[3] AND NOT FH_A_ST1_Done AND FH_Line0_Trigger_Ready_1 AND NOT FH_Line0_Error_Status_1;
FH_A_ST1_M[6] := _p9;
FH_A_ST1_OK := _p9;
(* Rung 6: NG判定 *)
_e10(CLK := FH_A_ST1_M[5] AND (FH_Line0_DINT_Result_Data_0_1 = (DINT#-1000)));
IF _e10.Q THEN
    HMI_MessageNo[0] := INT#114;
    Station_A_Data[1].Total_Judge := INT#9;
    Station_A_Data[1].Judgment_Details := INT#1;
END_IF;
_e11(CLK := FH_A_ST1_M[5] AND (FH_Line0_DINT_Result_Data_1_1 = (DINT#-1000)));
IF _e11.Q THEN
    HMI_MessageNo[0] := INT#115;
    Station_A_Data[1].Total_Judge := INT#9;
    Station_A_Data[1].Judgment_Details := INT#2;
END_IF;
_p12 := (_e10.Q OR _e11.Q OR FH_A_ST1_M[7]) AND NOT M9999 AND NOT Pause[3] AND NOT FH_A_ST1_Done AND FH_Line0_Trigger_Ready_1 AND NOT FH_Line0_Error_Status_1;
FH_A_ST1_M[7] := _p12;
FH_A_ST1_NG := _p12;

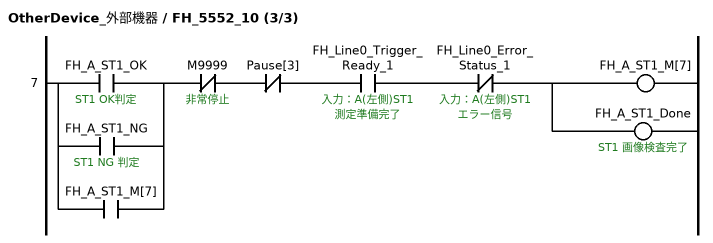
(* Rung 7 *)
_p13 := (FH_A_ST1_OK OR FH_A_ST1_NG OR FH_A_ST1_M[7]) AND NOT M9999 AND NOT Pause[3] AND FH_Line0_Trigger_Ready_1 AND NOT FH_Line0_Error_Status_1;
FH_A_ST1_M[7] := _p13;
FH_A_ST1_Done := _p13;

(* Section HMI: ladder, written here as Structured Text *)

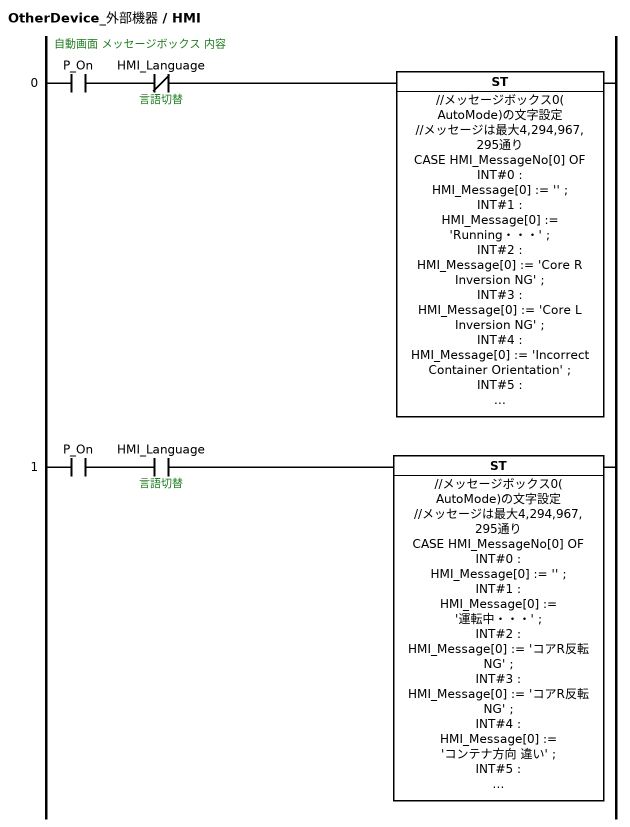
(* Rung 0: 自動画面 メッセージボックス 内容 *)
IF P_On AND NOT HMI_Language THEN
    //メッセージボックス0(AutoMode)の文字設定
    //メッセージは最大4,294,967,295通り
    	
    	CASE HMI_MessageNo[0] OF
    	
    	INT#0 :
    	HMI_Message[0] := '' ;
        INT#1 :
    	HMI_Message[0] := 'Running・・・' ;
    	INT#2 :
    	HMI_Message[0] := 'Core R Inversion NG' ;
    	INT#3 :
    	HMI_Message[0] := 'Core L Inversion NG' ;
    	INT#4 :
    	HMI_Message[0] := 'Incorrect Container Orientation' ;
    	INT#5 :
    	HMI_Message[0] := 'Packed Container Full' ;
         INT#6 :
    	HMI_Message[0] := 'No Container Added' ;
    	INT#7 :
    	HMI_Message[0] := 'Paused・・・' ;
        INT#8 :
    	HMI_Message[0] := 'R Stock Holder Qty Error' ;
    	INT#9 :
    	HMI_Message[0] := 'L Stock Holder Qty Error' ;
        INT#10 :
    	HMI_Message[0] := 'Step Running・・・' ;
    	INT#11 :
    	HMI_Message[0] := 'Work Discharge Complete' ;
    	INT#12 :
    	HMI_Message[0] := 'SD Error' ;
    	END_CASE;		
    	
END_IF;
(* Rung 1 *)
IF P_On AND HMI_Language THEN
    //メッセージボックス0(AutoMode)の文字設定
    //メッセージは最大4,294,967,295通り
    	
    	CASE HMI_MessageNo[0] OF
    	
    	INT#0 :
    	HMI_Message[0] := '' ;
    	INT#1 :
    	HMI_Message[0] := '運転中・・・' ;	
    	INT#2 :
    	HMI_Message[0] := 'コアR反転 NG' ;	
        INT#3 :
    	HMI_Message[0] := 'コアR反転 NG' ;
    	INT#4 :
    	HMI_Message[0] := 'コンテナ方向 違い' ;
    	INT#5 :
    	HMI_Message[0] := '梱包済みコンテナ 満杯 or 排出詰まり' ;
        INT#6 :
    	HMI_Message[0] := 'コンテナ 無 追加してください' ;
        INT#7 :
    	HMI_Message[0] := '一時停止中・・・' ;
        INT#8 :
    	HMI_Message[0] := '右ストックフォルダ 入数ミス 取り除いて 再スタート' ;
        INT#9 :
    	HMI_Message[0] := '左ストックフォルダ 入数ミス 取り除いて 再スタート' ;
    	INT#10 :
    	HMI_Message[0] := 'ステップ運転中・・・' ;
    	INT#11 :
    	HMI_Message[0] := 'ワーク排出完了' ;
    	INT#12 :
    	HMI_Message[0] := 'SDカードエラー' ;
    	END_CASE;		
    	
END_IF;
END_PROGRAM

